(* Logix 5000 project; controller TFF vendor 1 type 14 code 107 rev 33.11; software revision 33.04; part 5 of 38 *)

        [0,11].PID.KP := 0.1, [0,11].PID.KI := 0.1, [0,11].PID.BIAS := 23.09767, [0,11].PID.DB := 0.001, [0,11].PID.MAXO := 100.0, [0,11].PID.UPD := 0.25, [0,11].PID.ERR := 0.20000005, [0,11].PID.MAXCV := 100.0, [0,11].PID.MAXTIE := 100.0, [0,11].PID.DATA[0] := -23.098158, [0,11].PID.DATA[3] := 0.20000005, [0,11].PID.DATA[4] := 0.20000005, [0,11].PID.DATA[5] := 0.024420025, [0,11].PID.DATA[6] := 1.0, [0,11].PID.DATA[7] := 4.0, [0,11].PID.DATA[8] := 0.1, [0,11].PID.DATA[9] := 0.1, [0,11].PID.DATA[11] := 0.1, [0,11].PID.DATA[12] := 0.1, [0,11].PID.DATA[15] := 1.0, [0,11].PID.DATA[16] := 1.0, [0,13].RampTimer.PRE := 3600000, [0,13].StableTimer.PRE := 2000, [0,13].PIDTimer.PRE := 10000, [0,13].PIDTimer.EN := 1, [0,13].PIDTimer.TT := 1, [0,13].PID.CTL := 305173120, [0,13].PID.PVT := 1, [0,13].PID.CA := 1, [0,13].PID.NOBC := 1, [0,13].PID.NOZC := 1, [0,13].PID.INI := 1, [0,13].PID.OLH := 1, [0,13].PID.DVPA := 1, [0,13].PID.PVHA := 1, [0,13].PID.KP := 0.2, [0,13].PID.KI := 0.08, [0,13].PID.MAXS := 100.0, [0,13].PID.DB := 1.0, [0,13].PID.SO := 100.0, [0,13].PID.MAXO := 100.0, [0,13].PID.UPD := 0.01, [0,13].PID.PV := 43.925232, [0,13].PID.ERR := 43.925232, [0,13].PID.OUT := 100.0, [0,13].PID.MAXI := 100.0, [0,13].PID.TIE := 2.4420025, [0,13].PID.MAXCV := 100.0, [0,13].PID.MAXTIE := 4095.0, [0,13].PID.DATA[0] := 100.0, [0,13].PID.DATA[1] := 702.8037, [0,13].PID.DATA[2] := 43.925232, [0,13].PID.DATA[3] := 43.925232, [0,13].PID.DATA[5] := 1.0, [0,13].PID.DATA[6] := 1.0, [0,13].PID.DATA[7] := 0.16, [0,13].PID.DATA[8] := 0.2, [0,13].PID.DATA[9] := 0.08, [0,13].PID.DATA[11] := 0.2, [0,13].PID.DATA[12] := 0.08,
        [0,13].PID.DATA[15] := 1.0, [0,13].PID.DATA[16] := 0.024420025, [1,0].RampTimer.PRE := 3600000, [1,0].StableTimer.PRE := 5000, [1,0].PIDTimer.PRE := 250, [1,0].PIDTimer.ACC := 100, [1,0].PIDTimer.EN := 1, [1,0].PIDTimer.TT := 1, [1,0].PID.CTL := 25199488, [1,0].PID.MO := 1, [1,0].PID.PE := 1, [1,0].PID.INI := 1, [1,0].PID.DVPA := 1, [1,0].PID.PVLA := 1, [1,0].PID.PVHA := 1, [1,0].PID.SP := 66.66666, [1,0].PID.KP := 0.5, [1,0].PID.KI := 0.1, [1,0].PID.MAXS := 200.0, [1,0].PID.SO := 10.0, [1,0].PID.MAXO := 100.0, [1,0].PID.MINO := 10.0, [1,0].PID.UPD := 0.25, [1,0].PID.ERR := 66.66666, [1,0].PID.OUT := 10.0, [1,0].PID.MAXI := 200.0, [1,0].PID.TIE := 10.0, [1,0].PID.MAXCV := 100.0, [1,0].PID.MAXTIE := 100.0, [1,0].PID.DATA[0] := -6.666666, [1,0].PID.DATA[3] := 66.66666, [1,0].PID.DATA[4] := 66.66666, [1,0].PID.DATA[5] := 0.5, [1,0].PID.DATA[6] := 1.0, [1,0].PID.DATA[7] := 4.0, [1,0].PID.DATA[8] := 0.5, [1,0].PID.DATA[9] := 0.1, [1,0].PID.DATA[11] := 0.5, [1,0].PID.DATA[12] := 0.08333334, [1,0].PID.DATA[15] := 1.0, [1,0].PID.DATA[16] := 1.0, [1,1].Tag := 'FIC01', [1,1].Desc := 'Prim. Feed Pump Control', [1,1].LoopCfg := 1, [1,1].ManualEGU := '%', [1,1].Auto1EGU := 'LPM', [1,1].Auto2EGU := 'cm/h', [1,1].Manual := 1, [1,1].DBOK := 1, [1,1].RampEnable := 1, [1,1].PIDEnable := 1, [1,1].ManualOSR := 1, [1,1].RangeMax := 100.0, [1,1].RampRate := 5.0, [1,1].RampRateSave := 5.0, [1,1].Deadband := 5.0, [1,1].RampTimer.PRE := 3600000, [1,1].StableTimer.PRE := 10000, [1,1].StableTime := 10, [1,1].PIDTimer.PRE := 250,
        [1,1].CycleTimer.PRE := 2000, [1,1].PID.CTL := -2080340096, [1,1].PID.EN := 1, [1,1].PID.SWM := 1, [1,1].PID.INI := 1, [1,1].PID.DVNA := 1, [1,1].PID.DVPA := 1, [1,1].PID.PVLA := 1, [1,1].PID.PVHA := 1, [1,1].PID.KP := 0.7, [1,1].PID.KI := 1.4, [1,1].PID.KD := 0.013, [1,1].PID.MAXS := 22.0, [1,1].PID.DB := 0.001, [1,1].PID.MAXO := 100.0, [1,1].PID.UPD := 0.25, [1,1].PID.MAXI := 22.0, [1,1].PID.MAXCV := 100.0, [1,1].PID.MAXTIE := 22.0, [1,1].PID.DATA[5] := 4.5454545, [1,1].PID.DATA[6] := 1.0, [1,1].PID.DATA[7] := 4.013, [1,1].PID.DATA[8] := 0.7, [1,1].PID.DATA[9] := 1.4, [1,1].PID.DATA[10] := 0.013, [1,1].PID.DATA[11] := 0.7, [1,1].PID.DATA[12] := 1.4, [1,1].PID.DATA[13] := 0.013, [1,1].PID.DATA[15] := 1.0, [1,1].PID.DATA[16] := 4.5454545, [1,1].KP[0] := 700.0, [1,1].KI[0] := 1400.0, [1,1].KD[0] := 13.0, [1,1].Auto1Cfg := 1, [1,1].Auto2Cfg := 1, [1,1].Auto1PVCfg := 10, [1,1].Auto2PVCfg := 42, [1,1].Auto1RangeMax := 22.0, [1,1].Auto2RangeMax := 9999.0, [1,2].Tag := 'FIC02', [1,2].Desc := 'Sec. Feed Pump Control', [1,2].LoopCfg := 1, [1,2].ManualEGU := '%', [1,2].Auto1EGU := 'LPM', [1,2].Auto2EGU := 'cm/h', [1,2].Interlock := 1, [1,2].Manual := 1, [1,2].DBOK := 1, [1,2].RampEnable := 1, [1,2].PIDEnable := 1, [1,2].ManualOSR := 1, [1,2].RangeMax := 100.0, [1,2].RampRate := 5.0, [1,2].RampRateSave := 5.0, [1,2].Deadband := 5.0, [1,2].RampTimer.PRE := 3600000, [1,2].StableTimer.PRE := 10000, [1,2].StableTime := 10, [1,2].PIDTimer.PRE := 250, [1,2].CycleTimer.PRE := 2000,
        [1,2].PID.CTL := -2080340096, [1,2].PID.EN := 1, [1,2].PID.SWM := 1, [1,2].PID.INI := 1, [1,2].PID.DVNA := 1, [1,2].PID.DVPA := 1, [1,2].PID.PVLA := 1, [1,2].PID.PVHA := 1, [1,2].PID.KP := 0.7, [1,2].PID.KI := 1.4, [1,2].PID.KD := 0.013, [1,2].PID.MAXS := 22.0, [1,2].PID.DB := 0.001, [1,2].PID.MAXO := 100.0, [1,2].PID.UPD := 0.25, [1,2].PID.MAXI := 22.0, [1,2].PID.MAXCV := 100.0, [1,2].PID.MAXTIE := 100.0, [1,2].PID.DATA[5] := 4.5454545, [1,2].PID.DATA[6] := 1.0, [1,2].PID.DATA[7] := 4.013, [1,2].PID.DATA[8] := 0.7, [1,2].PID.DATA[9] := 1.4, [1,2].PID.DATA[10] := 0.013, [1,2].PID.DATA[11] := 0.7, [1,2].PID.DATA[12] := 1.4, [1,2].PID.DATA[13] := 0.013, [1,2].PID.DATA[15] := 1.0, [1,2].PID.DATA[16] := 1.0, [1,2].KP[0] := 700.0, [1,2].KI[0] := 1400.0, [1,2].KD[0] := 13.0, [1,2].DisOSR := 1, [1,2].Auto1Cfg := 1, [1,2].Auto2Cfg := 1, [1,2].Auto1PVCfg := 12, [1,2].Auto2PVCfg := 43, [1,2].Auto1RangeMax := 22.0, [1,2].Auto2RangeMax := 9999.0, [1,2].OutputAddress := 1, [1,3].Tag := 'PCV12', [1,3].Desc := 'Post Column PCV012 Control', [1,3].LoopCfg := 1, [1,3].ManualEGU := '%', [1,3].Enable := 1, [1,3].Manual := 1, [1,3].Stable := 1, [1,3].DBOK := 1, [1,3].Status := 3, [1,3].RampEnable := 1, [1,3].PIDEnable := 1, [1,3].ManualOSR := 1, [1,3].RangeMax := 100.0, [1,3].RampRate := 5.0, [1,3].RampRateSave := 5.0, [1,3].RampStart := 20.0, [1,3].RampTimer.PRE := 3600000, [1,3].StableTimer.PRE := 2300, [1,3].StableTimer.ACC := 2354, [1,3].StableTimer.EN := 1,
        [1,3].StableTimer.DN := 1, [1,3].PIDTimer.PRE := 250, [1,3].CycleTimer.PRE := 2000, [1,3].PID.CTL := -1946122368, [1,3].PID.EN := 1, [1,3].PID.DOE := 1, [1,3].PID.SWM := 1, [1,3].PID.INI := 1, [1,3].PID.DVNA := 1, [1,3].PID.DVPA := 1, [1,3].PID.PVLA := 1, [1,3].PID.PVHA := 1, [1,3].PID.KP := 0.001, [1,3].PID.KI := 0.001, [1,3].PID.BIAS := 30.796, [1,3].PID.MAXS := 4095.0, [1,3].PID.MAXO := 100.0, [1,3].PID.UPD := 0.01, [1,3].PID.MAXI := 4095.0, [1,3].PID.MAXCV := 100.0, [1,3].PID.MAXTIE := 100.0, [1,3].PID.DATA[0] := -30.796, [1,3].PID.DATA[5] := 0.024420025, [1,3].PID.DATA[6] := 1.0, [1,3].PID.DATA[7] := 0.16, [1,3].PID.DATA[8] := 0.001, [1,3].PID.DATA[9] := 0.001, [1,3].PID.DATA[11] := 0.001, [1,3].PID.DATA[12] := 0.001, [1,3].PID.DATA[15] := 1.0, [1,3].PID.DATA[16] := 1.0, [1,3].OutputAddress := 2, [1,4].Tag := 'PCV10', [1,4].Desc := 'Line Pump1 PCV010 Control', [1,4].ManualEGU := '%', [1,4].Manual := 1, [1,4].Status := 3, [1,4].RampEnable := 1, [1,4].PIDEnable := 1, [1,4].RangeMax := 100.0, [1,4].RampRate := 0.5, [1,4].RampRateSave := 0.5, [1,4].RampStart := 3.443, [1,4].RampTimer.PRE := 3600000, [1,4].StableTimer.PRE := 5000, [1,4].PIDTimer.PRE := 250, [1,4].CycleTimer.PRE := 2000, [1,4].PID.CTL := 35652992, [1,4].PID.CA := 1, [1,4].PID.NOBC := 1, [1,4].PID.DVNA := 1, [1,4].PID.PVLA := 1, [1,4].PID.PVHA := 1, [1,4].PID.SP := 19.6, [1,4].PID.KP := 0.1, [1,4].PID.KI := 0.3, [1,4].PID.MAXS := 150.0, [1,4].PID.MAXO := 100.0, [1,4].PID.UPD := 0.25, [1,4].PID.ERR := -19.6,
        [1,4].PID.MAXI := 150.0, [1,4].PID.MAXCV := 100.0, [1,4].PID.MAXTIE := 100.0, [1,4].PID.DATA[0] := 1.3066667, [1,4].PID.DATA[3] := -19.6, [1,4].PID.DATA[4] := 19.6, [1,4].PID.DATA[5] := 0.6666667, [1,4].PID.DATA[6] := 1.0, [1,4].PID.DATA[7] := 4.0, [1,4].PID.DATA[8] := 0.1, [1,4].PID.DATA[9] := 0.3, [1,4].PID.DATA[11] := 0.1, [1,4].PID.DATA[12] := 0.3, [1,4].PID.DATA[15] := 1.0, [1,4].PID.DATA[16] := 1.0, [1,4].OutputAddress := 2, [1,5].Tag := 'PCV11', [1,5].Desc := 'Line Pump2 PCV011 Control', [1,5].ManualEGU := '%', [1,5].Manual := 1, [1,5].Status := 3, [1,5].RampEnable := 1, [1,5].PIDEnable := 1, [1,5].RangeMax := 100.0, [1,5].RampRate := 0.5, [1,5].RampRateSave := 0.5, [1,5].RampStart := 4.417, [1,5].RampTimer.PRE := 3600000, [1,5].StableTimer.PRE := 1500, [1,5].PIDTimer.PRE := 250, [1,5].CycleTimer.PRE := 2000, [1,5].PID.CTL := 134218624, [1,5].PID.DOE := 1, [1,5].PID.DVPA := 1, [1,5].PID.PVLA := 1, [1,5].PID.PVHA := 1, [1,5].PID.SP := 350.0, [1,5].PID.KP := 40.0, [1,5].PID.KI := 0.5, [1,5].PID.BIAS := -847.4798, [1,5].PID.MAXS := 550.0, [1,5].PID.MAXO := 100.0, [1,5].PID.UPD := 0.25, [1,5].PID.ERR := 350.0, [1,5].PID.MAXI := 550.0, [1,5].PID.MAXCV := 100.0, [1,5].PID.MAXTIE := 100.0, [1,5].PID.DATA[0] := -1697.9749, [1,5].PID.DATA[1] := 1018.1818, [1,5].PID.DATA[3] := 350.0, [1,5].PID.DATA[4] := 350.0, [1,5].PID.DATA[5] := 0.18181819, [1,5].PID.DATA[6] := 1.0, [1,5].PID.DATA[7] := 4.0, [1,5].PID.DATA[8] := 40.0, [1,5].PID.DATA[9] := 0.5, [1,5].PID.DATA[11] := 40.0, [1,5].PID.DATA[12] := 0.5, [1,5].PID.DATA[15] := 1.0, [1,5].PID.DATA[16] := 1.0,
        [1,5].OutputAddress := 3, [1,6].StableTimer.PRE := 15000, [1,6].PIDTimer.EN := 1, [1,6].PIDTimer.TT := 1, [1,6].CycleTimer.PRE := 5000, [1,6].PID.CTL := 16810624, [1,6].PID.MO := 1, [1,6].PID.INI := 1, [1,6].PID.DVPA := 1, [1,6].PID.PVHA := 1, [1,6].PID.SP := 10.0, [1,6].PID.KP := 0.3, [1,6].PID.KI := 0.3, [1,6].PID.MAXS := 200.0, [1,6].PID.SO := 3.074094, [1,6].PID.MAXO := 100.0, [1,6].PID.UPD := 0.25, [1,6].PID.PV := 1.488363, [1,6].PID.ERR := 8.511638, [1,6].PID.OUT := 3.074094, [1,6].PID.MAXI := 200.0, [1,6].PID.TIE := 3.074094, [1,6].PID.MAXCV := 200.0, [1,6].PID.MAXTIE := 200.0, [1,6].PID.DATA[0] := 1.797348, [1,6].PID.DATA[1] := -11.9069, [1,6].PID.DATA[2] := 1.488363, [1,6].PID.DATA[3] := 8.511638, [1,6].PID.DATA[4] := 10.0, [1,6].PID.DATA[5] := 0.5, [1,6].PID.DATA[6] := 1.0, [1,6].PID.DATA[7] := 4.0, [1,6].PID.DATA[8] := 0.3, [1,6].PID.DATA[9] := 0.3, [1,6].PID.DATA[11] := 0.3, [1,6].PID.DATA[12] := 0.3, [1,6].PID.DATA[15] := 2.0, [1,6].PID.DATA[16] := 0.5, [1,7].StableTimer.PRE := 200, [1,7].PIDTimer.PRE := 250, [1,7].PIDTimer.EN := 1, [1,7].PIDTimer.TT := 1, [1,7].CycleTimer.PRE := 10000, [1,7].PID.CTL := 16810880, [1,7].PID.MO := 1, [1,7].PID.INI := 1, [1,7].PID.DVPA := 1, [1,7].PID.PVLA := 1, [1,7].PID.PVHA := 1, [1,7].PID.SP := 10.0, [1,7].PID.KP := 2.0, [1,7].PID.KI := 0.2, [1,7].PID.KD := 0.3, [1,7].PID.BIAS := 50.0, [1,7].PID.DB := 0.01, [1,7].PID.SO := 80.0, [1,7].PID.MAXO := 100.0, [1,7].PID.UPD := 0.25, [1,7].PID.ERR := 10.0, [1,7].PID.OUT := 80.0,
        [1,7].PID.TIE := 80.0, [1,7].PID.MAXCV := 100.0, [1,7].PID.MAXTIE := 100.0, [1,7].PID.DATA[0] := 29.511597, [1,7].PID.DATA[3] := 10.0, [1,7].PID.DATA[4] := 10.0, [1,7].PID.DATA[5] := 0.024420025, [1,7].PID.DATA[6] := 1.0, [1,7].PID.DATA[7] := 4.3, [1,7].PID.DATA[8] := 2.0, [1,7].PID.DATA[9] := 0.2, [1,7].PID.DATA[10] := 0.3, [1,7].PID.DATA[11] := 2.0, [1,7].PID.DATA[12] := 0.2, [1,7].PID.DATA[13] := 0.3, [1,7].PID.DATA[15] := 1.0, [1,7].PID.DATA[16] := 1.0, [1,8].StableTimer.PRE := 15000, [1,8].PIDTimer.PRE := 250, [1,8].CycleTimer.PRE := 20000, [1,8].PID.CTL := 33555584, [1,8].PID.CA := 1, [1,8].PID.DVNA := 1, [1,8].PID.PVHA := 1, [1,8].PID.SP := 27.0, [1,8].PID.KP := 1.0, [1,8].PID.KI := 0.1, [1,8].PID.MAXS := 100.0, [1,8].PID.MAXO := 100.0, [1,8].PID.UPD := 0.25, [1,8].PID.PV := 18.2328, [1,8].PID.ERR := -8.767202, [1,8].PID.MAXI := 100.0, [1,8].PID.MAXCV := 100.0, [1,8].PID.MAXTIE := 100.0, [1,8].PID.DATA[0] := 8.767202, [1,8].PID.DATA[1] := 291.7248, [1,8].PID.DATA[2] := 18.2328, [1,8].PID.DATA[3] := -8.767202, [1,8].PID.DATA[4] := 27.0, [1,8].PID.DATA[5] := 1.0, [1,8].PID.DATA[6] := 1.0, [1,8].PID.DATA[7] := 4.0, [1,8].PID.DATA[8] := 1.0, [1,8].PID.DATA[9] := 0.1, [1,8].PID.DATA[11] := 1.0, [1,8].PID.DATA[12] := 0.1, [1,8].PID.DATA[15] := 1.0, [1,8].PID.DATA[16] := 1.0, [1,11].RampTimer.PRE := 100000, [1,11].StableTimer.PRE := 200, [1,11].PIDTimer.PRE := 250, [1,11].PIDTimer.ACC := 230, [1,11].PIDTimer.EN := 1, [1,11].PIDTimer.TT := 1, [1,11].PID.CTL := 67142528, [1,11].PID.SWM := 1, [1,11].PID.INI := 1, [1,11].PID.DVPA := 1, [1,11].PID.PVLA := 1,
        [1,11].PID.PVHA := 1, [1,11].PID.SP := 0.20000005, [1,11].PID.KP := 0.1, [1,11].PID.KI := 0.1, [1,11].PID.BIAS := 23.09767, [1,11].PID.DB := 0.001, [1,11].PID.MAXO := 100.0, [1,11].PID.UPD := 0.25, [1,11].PID.ERR := 0.20000005, [1,11].PID.MAXCV := 100.0, [1,11].PID.MAXTIE := 100.0, [1,11].PID.DATA[0] := -23.098158, [1,11].PID.DATA[3] := 0.20000005, [1,11].PID.DATA[4] := 0.20000005, [1,11].PID.DATA[5] := 0.024420025, [1,11].PID.DATA[6] := 1.0, [1,11].PID.DATA[7] := 4.0, [1,11].PID.DATA[8] := 0.1, [1,11].PID.DATA[9] := 0.1, [1,11].PID.DATA[11] := 0.1, [1,11].PID.DATA[12] := 0.1, [1,11].PID.DATA[15] := 1.0, [1,11].PID.DATA[16] := 1.0, [1,13].RampTimer.PRE := 3600000, [1,13].StableTimer.PRE := 2000, [1,13].PIDTimer.PRE := 10000, [1,13].PIDTimer.EN := 1, [1,13].PIDTimer.TT := 1, [1,13].PID.CTL := 305173120, [1,13].PID.PVT := 1, [1,13].PID.CA := 1, [1,13].PID.NOBC := 1, [1,13].PID.NOZC := 1, [1,13].PID.INI := 1, [1,13].PID.OLH := 1, [1,13].PID.DVPA := 1, [1,13].PID.PVHA := 1, [1,13].PID.KP := 0.2, [1,13].PID.KI := 0.08, [1,13].PID.MAXS := 100.0, [1,13].PID.DB := 1.0, [1,13].PID.SO := 100.0, [1,13].PID.MAXO := 100.0, [1,13].PID.UPD := 0.01, [1,13].PID.PV := 43.925232, [1,13].PID.ERR := 43.925232, [1,13].PID.OUT := 100.0, [1,13].PID.MAXI := 100.0, [1,13].PID.TIE := 2.4420025, [1,13].PID.MAXCV := 100.0, [1,13].PID.MAXTIE := 4095.0, [1,13].PID.DATA[0] := 100.0, [1,13].PID.DATA[1] := 702.8037, [1,13].PID.DATA[2] := 43.925232, [1,13].PID.DATA[3] := 43.925232, [1,13].PID.DATA[5] := 1.0, [1,13].PID.DATA[6] := 1.0, [1,13].PID.DATA[7] := 0.16, [1,13].PID.DATA[8] := 0.2, [1,13].PID.DATA[9] := 0.08,
        [1,13].PID.DATA[11] := 0.2, [1,13].PID.DATA[12] := 0.08, [1,13].PID.DATA[15] := 1.0, [1,13].PID.DATA[16] := 0.024420025, [2,0].RampTimer.PRE := 3600000, [2,0].StableTimer.PRE := 5000, [2,0].PIDTimer.PRE := 250, [2,0].PIDTimer.ACC := 100, [2,0].PIDTimer.EN := 1, [2,0].PIDTimer.TT := 1, [2,0].PID.CTL := 25199488, [2,0].PID.MO := 1, [2,0].PID.PE := 1, [2,0].PID.INI := 1, [2,0].PID.DVPA := 1, [2,0].PID.PVLA := 1, [2,0].PID.PVHA := 1, [2,0].PID.SP := 66.66666, [2,0].PID.KP := 0.5, [2,0].PID.KI := 0.1, [2,0].PID.MAXS := 200.0, [2,0].PID.SO := 10.0, [2,0].PID.MAXO := 100.0, [2,0].PID.MINO := 10.0, [2,0].PID.UPD := 0.25, [2,0].PID.ERR := 66.66666, [2,0].PID.OUT := 10.0, [2,0].PID.MAXI := 200.0, [2,0].PID.TIE := 10.0, [2,0].PID.MAXCV := 100.0, [2,0].PID.MAXTIE := 100.0, [2,0].PID.DATA[0] := -6.666666, [2,0].PID.DATA[3] := 66.66666, [2,0].PID.DATA[4] := 66.66666, [2,0].PID.DATA[5] := 0.5, [2,0].PID.DATA[6] := 1.0, [2,0].PID.DATA[7] := 4.0, [2,0].PID.DATA[8] := 0.5, [2,0].PID.DATA[9] := 0.1, [2,0].PID.DATA[11] := 0.5, [2,0].PID.DATA[12] := 0.08333334, [2,0].PID.DATA[15] := 1.0, [2,0].PID.DATA[16] := 1.0, [2,1].Tag := 'FIC01', [2,1].Desc := 'Prim. Feed Pump Control', [2,1].LoopCfg := 1, [2,1].ManualEGU := '%', [2,1].Auto1EGU := 'LPM', [2,1].Auto2EGU := 'cm/h', [2,1].Manual := 1, [2,1].DBOK := 1, [2,1].RampEnable := 1, [2,1].PIDEnable := 1, [2,1].ManualOSR := 1, [2,1].RangeMax := 100.0, [2,1].RampRate := 5.0, [2,1].RampRateSave := 5.0, [2,1].Deadband := 5.0, [2,1].RampTimer.PRE := 3600000, [2,1].StableTimer.PRE := 10000,
        [2,1].StableTime := 10, [2,1].PIDTimer.PRE := 250, [2,1].CycleTimer.PRE := 2000, [2,1].PID.CTL := -2080340096, [2,1].PID.EN := 1, [2,1].PID.SWM := 1, [2,1].PID.INI := 1, [2,1].PID.DVNA := 1, [2,1].PID.DVPA := 1, [2,1].PID.PVLA := 1, [2,1].PID.PVHA := 1, [2,1].PID.KP := 0.7, [2,1].PID.KI := 1.4, [2,1].PID.KD := 0.013, [2,1].PID.MAXS := 22.0, [2,1].PID.DB := 0.001, [2,1].PID.MAXO := 100.0, [2,1].PID.UPD := 0.25, [2,1].PID.MAXI := 22.0, [2,1].PID.MAXCV := 100.0, [2,1].PID.MAXTIE := 22.0, [2,1].PID.DATA[5] := 4.5454545, [2,1].PID.DATA[6] := 1.0, [2,1].PID.DATA[7] := 4.013, [2,1].PID.DATA[8] := 0.7, [2,1].PID.DATA[9] := 1.4, [2,1].PID.DATA[10] := 0.013, [2,1].PID.DATA[11] := 0.7, [2,1].PID.DATA[12] := 1.4, [2,1].PID.DATA[13] := 0.013, [2,1].PID.DATA[15] := 1.0, [2,1].PID.DATA[16] := 4.5454545, [2,1].KP[0] := 700.0, [2,1].KI[0] := 1400.0, [2,1].KD[0] := 13.0, [2,1].Auto1Cfg := 1, [2,1].Auto2Cfg := 1, [2,1].Auto1PVCfg := 10, [2,1].Auto2PVCfg := 42, [2,1].Auto1RangeMax := 22.0, [2,1].Auto2RangeMax := 9999.0, [2,2].Tag := 'FIC02', [2,2].Desc := 'Sec. Feed Pump Control', [2,2].LoopCfg := 1, [2,2].ManualEGU := '%', [2,2].Auto1EGU := 'LPM', [2,2].Auto2EGU := 'cm/h', [2,2].Interlock := 1, [2,2].Manual := 1, [2,2].DBOK := 1, [2,2].RampEnable := 1, [2,2].PIDEnable := 1, [2,2].ManualOSR := 1, [2,2].RangeMax := 100.0, [2,2].RampRate := 5.0, [2,2].RampRateSave := 5.0, [2,2].Deadband := 5.0, [2,2].RampTimer.PRE := 3600000, [2,2].StableTimer.PRE := 10000, [2,2].StableTime := 10,
        [2,2].PIDTimer.PRE := 250, [2,2].CycleTimer.PRE := 2000, [2,2].PID.CTL := -2080340096, [2,2].PID.EN := 1, [2,2].PID.SWM := 1, [2,2].PID.INI := 1, [2,2].PID.DVNA := 1, [2,2].PID.DVPA := 1, [2,2].PID.PVLA := 1, [2,2].PID.PVHA := 1, [2,2].PID.KP := 0.7, [2,2].PID.KI := 1.4, [2,2].PID.KD := 0.013, [2,2].PID.MAXS := 22.0, [2,2].PID.DB := 0.001, [2,2].PID.MAXO := 100.0, [2,2].PID.UPD := 0.25, [2,2].PID.MAXI := 22.0, [2,2].PID.MAXCV := 100.0, [2,2].PID.MAXTIE := 100.0, [2,2].PID.DATA[5] := 4.5454545, [2,2].PID.DATA[6] := 1.0, [2,2].PID.DATA[7] := 4.013, [2,2].PID.DATA[8] := 0.7, [2,2].PID.DATA[9] := 1.4, [2,2].PID.DATA[10] := 0.013, [2,2].PID.DATA[11] := 0.7, [2,2].PID.DATA[12] := 1.4, [2,2].PID.DATA[13] := 0.013, [2,2].PID.DATA[15] := 1.0, [2,2].PID.DATA[16] := 1.0, [2,2].KP[0] := 700.0, [2,2].KI[0] := 1400.0, [2,2].KD[0] := 13.0, [2,2].DisOSR := 1, [2,2].Auto1Cfg := 1, [2,2].Auto2Cfg := 1, [2,2].Auto1PVCfg := 12, [2,2].Auto2PVCfg := 43, [2,2].Auto1RangeMax := 22.0, [2,2].Auto2RangeMax := 9999.0, [2,2].OutputAddress := 1, [2,3].Tag := 'PCV12', [2,3].Desc := 'Post Column PCV012 Control', [2,3].LoopCfg := 1, [2,3].ManualEGU := '%', [2,3].Enable := 1, [2,3].Manual := 1, [2,3].Stable := 1, [2,3].DBOK := 1, [2,3].Status := 3, [2,3].RampEnable := 1, [2,3].PIDEnable := 1, [2,3].ManualOSR := 1, [2,3].RangeMax := 100.0, [2,3].RampRate := 5.0, [2,3].RampRateSave := 5.0, [2,3].RampStart := 20.0, [2,3].RampTimer.PRE := 3600000, [2,3].StableTimer.PRE := 2300,
        [2,3].StableTimer.ACC := 2354, [2,3].StableTimer.EN := 1, [2,3].StableTimer.DN := 1, [2,3].PIDTimer.PRE := 250, [2,3].CycleTimer.PRE := 2000, [2,3].PID.CTL := -1946122368, [2,3].PID.EN := 1, [2,3].PID.DOE := 1, [2,3].PID.SWM := 1, [2,3].PID.INI := 1, [2,3].PID.DVNA := 1, [2,3].PID.DVPA := 1, [2,3].PID.PVLA := 1, [2,3].PID.PVHA := 1, [2,3].PID.KP := 0.001, [2,3].PID.KI := 0.001, [2,3].PID.BIAS := 30.796, [2,3].PID.MAXS := 4095.0, [2,3].PID.MAXO := 100.0, [2,3].PID.UPD := 0.01, [2,3].PID.MAXI := 4095.0, [2,3].PID.MAXCV := 100.0, [2,3].PID.MAXTIE := 100.0, [2,3].PID.DATA[0] := -30.796, [2,3].PID.DATA[5] := 0.024420025, [2,3].PID.DATA[6] := 1.0, [2,3].PID.DATA[7] := 0.16, [2,3].PID.DATA[8] := 0.001, [2,3].PID.DATA[9] := 0.001, [2,3].PID.DATA[11] := 0.001, [2,3].PID.DATA[12] := 0.001, [2,3].PID.DATA[15] := 1.0, [2,3].PID.DATA[16] := 1.0, [2,3].OutputAddress := 2, [2,4].Tag := 'PCV10', [2,4].Desc := 'Line Pump1 PCV010 Control', [2,4].ManualEGU := '%', [2,4].Manual := 1, [2,4].Status := 3, [2,4].RampEnable := 1, [2,4].PIDEnable := 1, [2,4].RangeMax := 100.0, [2,4].RampRate := 0.5, [2,4].RampRateSave := 0.5, [2,4].RampStart := 3.443, [2,4].RampTimer.PRE := 3600000, [2,4].StableTimer.PRE := 5000, [2,4].PIDTimer.PRE := 250, [2,4].CycleTimer.PRE := 2000, [2,4].PID.CTL := 35652992, [2,4].PID.CA := 1, [2,4].PID.NOBC := 1, [2,4].PID.DVNA := 1, [2,4].PID.PVLA := 1, [2,4].PID.PVHA := 1, [2,4].PID.SP := 19.6, [2,4].PID.KP := 0.1, [2,4].PID.KI := 0.3, [2,4].PID.MAXS := 150.0, [2,4].PID.MAXO := 100.0,
        [2,4].PID.UPD := 0.25, [2,4].PID.ERR := -19.6, [2,4].PID.MAXI := 150.0, [2,4].PID.MAXCV := 100.0, [2,4].PID.MAXTIE := 100.0, [2,4].PID.DATA[0] := 1.3066667, [2,4].PID.DATA[3] := -19.6, [2,4].PID.DATA[4] := 19.6, [2,4].PID.DATA[5] := 0.6666667, [2,4].PID.DATA[6] := 1.0, [2,4].PID.DATA[7] := 4.0, [2,4].PID.DATA[8] := 0.1, [2,4].PID.DATA[9] := 0.3, [2,4].PID.DATA[11] := 0.1, [2,4].PID.DATA[12] := 0.3, [2,4].PID.DATA[15] := 1.0, [2,4].PID.DATA[16] := 1.0, [2,4].OutputAddress := 2, [2,5].Tag := 'PCV11', [2,5].Desc := 'Line Pump2 PCV011 Control', [2,5].ManualEGU := '%', [2,5].Manual := 1, [2,5].Status := 3, [2,5].RampEnable := 1, [2,5].PIDEnable := 1, [2,5].RangeMax := 100.0, [2,5].RampRate := 0.5, [2,5].RampRateSave := 0.5, [2,5].RampStart := 4.417, [2,5].RampTimer.PRE := 3600000, [2,5].StableTimer.PRE := 1500, [2,5].PIDTimer.PRE := 250, [2,5].CycleTimer.PRE := 2000, [2,5].PID.CTL := 134218624, [2,5].PID.DOE := 1, [2,5].PID.DVPA := 1, [2,5].PID.PVLA := 1, [2,5].PID.PVHA := 1, [2,5].PID.SP := 350.0, [2,5].PID.KP := 40.0, [2,5].PID.KI := 0.5, [2,5].PID.BIAS := -847.4798, [2,5].PID.MAXS := 550.0, [2,5].PID.MAXO := 100.0, [2,5].PID.UPD := 0.25, [2,5].PID.ERR := 350.0, [2,5].PID.MAXI := 550.0, [2,5].PID.MAXCV := 100.0, [2,5].PID.MAXTIE := 100.0, [2,5].PID.DATA[0] := -1697.9749, [2,5].PID.DATA[1] := 1018.1818, [2,5].PID.DATA[3] := 350.0, [2,5].PID.DATA[4] := 350.0, [2,5].PID.DATA[5] := 0.18181819, [2,5].PID.DATA[6] := 1.0, [2,5].PID.DATA[7] := 4.0, [2,5].PID.DATA[8] := 40.0, [2,5].PID.DATA[9] := 0.5, [2,5].PID.DATA[11] := 40.0, [2,5].PID.DATA[12] := 0.5,
        [2,5].PID.DATA[15] := 1.0, [2,5].PID.DATA[16] := 1.0, [2,5].OutputAddress := 3, [2,6].StableTimer.PRE := 15000, [2,6].PIDTimer.EN := 1, [2,6].PIDTimer.TT := 1, [2,6].CycleTimer.PRE := 5000, [2,6].PID.CTL := 16810624, [2,6].PID.MO := 1, [2,6].PID.INI := 1, [2,6].PID.DVPA := 1, [2,6].PID.PVHA := 1, [2,6].PID.SP := 10.0, [2,6].PID.KP := 0.3, [2,6].PID.KI := 0.3, [2,6].PID.MAXS := 200.0, [2,6].PID.SO := 3.074094, [2,6].PID.MAXO := 100.0, [2,6].PID.UPD := 0.25, [2,6].PID.PV := 1.488363, [2,6].PID.ERR := 8.511638, [2,6].PID.OUT := 3.074094, [2,6].PID.MAXI := 200.0, [2,6].PID.TIE := 3.074094, [2,6].PID.MAXCV := 200.0, [2,6].PID.MAXTIE := 200.0, [2,6].PID.DATA[0] := 1.797348, [2,6].PID.DATA[1] := -11.9069, [2,6].PID.DATA[2] := 1.488363, [2,6].PID.DATA[3] := 8.511638, [2,6].PID.DATA[4] := 10.0, [2,6].PID.DATA[5] := 0.5, [2,6].PID.DATA[6] := 1.0, [2,6].PID.DATA[7] := 4.0, [2,6].PID.DATA[8] := 0.3, [2,6].PID.DATA[9] := 0.3, [2,6].PID.DATA[11] := 0.3, [2,6].PID.DATA[12] := 0.3, [2,6].PID.DATA[15] := 2.0, [2,6].PID.DATA[16] := 0.5, [2,7].StableTimer.PRE := 200, [2,7].PIDTimer.PRE := 250, [2,7].PIDTimer.EN := 1, [2,7].PIDTimer.TT := 1, [2,7].CycleTimer.PRE := 10000, [2,7].PID.CTL := 16810880, [2,7].PID.MO := 1, [2,7].PID.INI := 1, [2,7].PID.DVPA := 1, [2,7].PID.PVLA := 1, [2,7].PID.PVHA := 1, [2,7].PID.SP := 10.0, [2,7].PID.KP := 2.0, [2,7].PID.KI := 0.2, [2,7].PID.KD := 0.3, [2,7].PID.BIAS := 50.0, [2,7].PID.DB := 0.01, [2,7].PID.SO := 80.0, [2,7].PID.MAXO := 100.0, [2,7].PID.UPD := 0.25,
        [2,7].PID.ERR := 10.0, [2,7].PID.OUT := 80.0, [2,7].PID.TIE := 80.0, [2,7].PID.MAXCV := 100.0, [2,7].PID.MAXTIE := 100.0, [2,7].PID.DATA[0] := 29.511597, [2,7].PID.DATA[3] := 10.0, [2,7].PID.DATA[4] := 10.0, [2,7].PID.DATA[5] := 0.024420025, [2,7].PID.DATA[6] := 1.0, [2,7].PID.DATA[7] := 4.3, [2,7].PID.DATA[8] := 2.0, [2,7].PID.DATA[9] := 0.2, [2,7].PID.DATA[10] := 0.3, [2,7].PID.DATA[11] := 2.0, [2,7].PID.DATA[12] := 0.2, [2,7].PID.DATA[13] := 0.3, [2,7].PID.DATA[15] := 1.0, [2,7].PID.DATA[16] := 1.0, [2,8].StableTimer.PRE := 15000, [2,8].PIDTimer.PRE := 250, [2,8].CycleTimer.PRE := 20000, [2,8].PID.CTL := 33555584, [2,8].PID.CA := 1, [2,8].PID.DVNA := 1, [2,8].PID.PVHA := 1, [2,8].PID.SP := 27.0, [2,8].PID.KP := 1.0, [2,8].PID.KI := 0.1, [2,8].PID.MAXS := 100.0, [2,8].PID.MAXO := 100.0, [2,8].PID.UPD := 0.25, [2,8].PID.PV := 18.2328, [2,8].PID.ERR := -8.767202, [2,8].PID.MAXI := 100.0, [2,8].PID.MAXCV := 100.0, [2,8].PID.MAXTIE := 100.0, [2,8].PID.DATA[0] := 8.767202, [2,8].PID.DATA[1] := 291.7248, [2,8].PID.DATA[2] := 18.2328, [2,8].PID.DATA[3] := -8.767202, [2,8].PID.DATA[4] := 27.0, [2,8].PID.DATA[5] := 1.0, [2,8].PID.DATA[6] := 1.0, [2,8].PID.DATA[7] := 4.0, [2,8].PID.DATA[8] := 1.0, [2,8].PID.DATA[9] := 0.1, [2,8].PID.DATA[11] := 1.0, [2,8].PID.DATA[12] := 0.1, [2,8].PID.DATA[15] := 1.0, [2,8].PID.DATA[16] := 1.0, [2,11].RampTimer.PRE := 100000, [2,11].StableTimer.PRE := 200, [2,11].PIDTimer.PRE := 250, [2,11].PIDTimer.ACC := 230, [2,11].PIDTimer.EN := 1, [2,11].PIDTimer.TT := 1, [2,11].PID.CTL := 67142528, [2,11].PID.SWM := 1, [2,11].PID.INI := 1,
        [2,11].PID.DVPA := 1, [2,11].PID.PVLA := 1, [2,11].PID.PVHA := 1, [2,11].PID.SP := 0.20000005, [2,11].PID.KP := 0.1, [2,11].PID.KI := 0.1, [2,11].PID.BIAS := 23.09767, [2,11].PID.DB := 0.001, [2,11].PID.MAXO := 100.0, [2,11].PID.UPD := 0.25, [2,11].PID.ERR := 0.20000005, [2,11].PID.MAXCV := 100.0, [2,11].PID.MAXTIE := 100.0, [2,11].PID.DATA[0] := -23.098158, [2,11].PID.DATA[3] := 0.20000005, [2,11].PID.DATA[4] := 0.20000005, [2,11].PID.DATA[5] := 0.024420025, [2,11].PID.DATA[6] := 1.0, [2,11].PID.DATA[7] := 4.0, [2,11].PID.DATA[8] := 0.1, [2,11].PID.DATA[9] := 0.1, [2,11].PID.DATA[11] := 0.1, [2,11].PID.DATA[12] := 0.1, [2,11].PID.DATA[15] := 1.0, [2,11].PID.DATA[16] := 1.0, [2,13].RampTimer.PRE := 3600000, [2,13].StableTimer.PRE := 2000, [2,13].PIDTimer.PRE := 10000, [2,13].PIDTimer.EN := 1, [2,13].PIDTimer.TT := 1, [2,13].PID.CTL := 305173120, [2,13].PID.PVT := 1, [2,13].PID.CA := 1, [2,13].PID.NOBC := 1, [2,13].PID.NOZC := 1, [2,13].PID.INI := 1, [2,13].PID.OLH := 1, [2,13].PID.DVPA := 1, [2,13].PID.PVHA := 1, [2,13].PID.KP := 0.2, [2,13].PID.KI := 0.08, [2,13].PID.MAXS := 100.0, [2,13].PID.DB := 1.0, [2,13].PID.SO := 100.0, [2,13].PID.MAXO := 100.0, [2,13].PID.UPD := 0.01, [2,13].PID.PV := 43.925232, [2,13].PID.ERR := 43.925232, [2,13].PID.OUT := 100.0, [2,13].PID.MAXI := 100.0, [2,13].PID.TIE := 2.4420025, [2,13].PID.MAXCV := 100.0, [2,13].PID.MAXTIE := 4095.0, [2,13].PID.DATA[0] := 100.0, [2,13].PID.DATA[1] := 702.8037, [2,13].PID.DATA[2] := 43.925232, [2,13].PID.DATA[3] := 43.925232, [2,13].PID.DATA[5] := 1.0, [2,13].PID.DATA[6] := 1.0, [2,13].PID.DATA[7] := 0.16,
        [2,13].PID.DATA[8] := 0.2, [2,13].PID.DATA[9] := 0.08, [2,13].PID.DATA[11] := 0.2, [2,13].PID.DATA[12] := 0.08, [2,13].PID.DATA[15] := 1.0, [2,13].PID.DATA[16] := 0.024420025, [3,1].LoopCfg := 1, [3,1].DBOK := 1, [3,1].RampEnable := 1, [3,1].PIDEnable := 1, [3,1].RangeMax := 100.0, [3,1].RampRate := 0.5, [3,1].RampRateSave := 0.5, [3,1].RampTimer.PRE := 3600000, [3,1].PIDTimer.PRE := 250, [3,1].PIDTimer.EN := 1, [3,1].PIDTimer.TT := 1, [3,1].CycleTimer.PRE := 2000, [3,1].PID.CTL := 67108864, [3,1].PID.SWM := 1, [3,1].PID.MAXS := 25.0, [3,1].PID.MAXO := 100.0, [3,1].PID.MAXI := 25.0, [3,1].PID.MAXCV := 100.0, [3,1].PID.MAXTIE := 25.0, [3,1].PID.DATA[5] := 4.0, [3,1].PID.DATA[6] := 1.0, [3,1].PID.DATA[15] := 1.0, [3,1].PID.DATA[16] := 4.0, [3,1].Auto1Cfg := 1, [3,1].Auto2Cfg := 1, [3,1].Auto1PVCfg := 10, [3,1].Auto2PVCfg := 42, [3,1].Auto1RangeMax := 55.0, [3,2].LoopCfg := 1, [3,2].DBOK := 1, [3,2].RampEnable := 1, [3,2].PIDEnable := 1, [3,2].RangeMax := 100.0, [3,2].RampRate := 0.5, [3,2].RampRateSave := 0.5, [3,2].RampTimer.PRE := 3600000, [3,2].PIDTimer.PRE := 250, [3,2].PIDTimer.EN := 1, [3,2].PIDTimer.TT := 1, [3,2].CycleTimer.PRE := 2000, [3,2].PID.CTL := 67108864, [3,2].PID.SWM := 1, [3,2].PID.MAXO := 100.0, [3,2].PID.MAXCV := 100.0, [3,2].PID.MAXTIE := 100.0, [3,2].PID.DATA[5] := 0.024420025, [3,2].PID.DATA[6] := 1.0, [3,2].PID.DATA[15] := 1.0, [3,2].PID.DATA[16] := 1.0, [3,2].Auto1Cfg := 1, [3,2].Auto2Cfg := 1, [3,2].Auto1PVCfg := 12, [3,2].Auto2PVCfg := 43, [3,2].Auto1RangeMax := 30.0,
        [3,2].OutputAddress := 1, [3,3].LoopCfg := 1, [3,3].Enable := 1, [3,3].Manual := 1, [3,3].Status := 9, [3,3].RampEnable := 1, [3,3].PIDEnable := 1, [3,3].RangeMax := 100.0, [3,3].RampRate := 0.5, [3,3].RampRateSave := 0.5, [3,3].RampTimer.PRE := 3600000, [3,3].PIDTimer.PRE := 250, [3,3].PIDTimer.EN := 1, [3,3].PIDTimer.TT := 1, [3,3].CycleTimer.PRE := 2000, [3,3].PID.CTL := 67108864, [3,3].PID.SWM := 1, [3,3].PID.MAXS := 4095.0, [3,3].PID.MAXO := 100.0, [3,3].PID.MAXI := 4095.0, [3,3].PID.MAXCV := 100.0, [3,3].PID.MAXTIE := 100.0, [3,3].PID.DATA[5] := 0.024420025, [3,3].PID.DATA[6] := 1.0, [3,3].PID.DATA[15] := 1.0, [3,3].PID.DATA[16] := 1.0, [3,3].OutputAddress := 2, [4,0].RampTimer.PRE := 3600000, [4,0].StableTimer.PRE := 5000, [4,0].PIDTimer.PRE := 250, [4,0].PIDTimer.ACC := 100, [4,0].PIDTimer.EN := 1, [4,0].PIDTimer.TT := 1, [4,0].PID.CTL := 25199488, [4,0].PID.MO := 1, [4,0].PID.PE := 1, [4,0].PID.INI := 1, [4,0].PID.DVPA := 1, [4,0].PID.PVLA := 1, [4,0].PID.PVHA := 1, [4,0].PID.SP := 66.66666, [4,0].PID.KP := 0.5, [4,0].PID.KI := 0.1, [4,0].PID.MAXS := 200.0, [4,0].PID.SO := 10.0, [4,0].PID.MAXO := 100.0, [4,0].PID.MINO := 10.0, [4,0].PID.UPD := 0.25, [4,0].PID.ERR := 66.66666, [4,0].PID.OUT := 10.0, [4,0].PID.MAXI := 200.0, [4,0].PID.TIE := 10.0, [4,0].PID.MAXCV := 100.0, [4,0].PID.MAXTIE := 100.0, [4,0].PID.DATA[0] := -6.666666, [4,0].PID.DATA[3] := 66.66666, [4,0].PID.DATA[4] := 66.66666, [4,0].PID.DATA[5] := 0.5, [4,0].PID.DATA[6] := 1.0, [4,0].PID.DATA[7] := 4.0,
        [4,0].PID.DATA[8] := 0.5, [4,0].PID.DATA[9] := 0.1, [4,0].PID.DATA[11] := 0.5, [4,0].PID.DATA[12] := 0.08333334, [4,0].PID.DATA[15] := 1.0, [4,0].PID.DATA[16] := 1.0, [4,1].Tag := 'FIC01', [4,1].Desc := 'Prim. Feed Pump Control', [4,1].LoopCfg := 1, [4,1].ManualEGU := '%', [4,1].Auto1EGU := 'LPM', [4,1].Auto2EGU := 'cm/h', [4,1].Manual := 1, [4,1].DBOK := 1, [4,1].RampEnable := 1, [4,1].PIDEnable := 1, [4,1].ManualOSR := 1, [4,1].PVAuto2 := 2400.0, [4,1].RangeMax := 100.0, [4,1].RampRate := 5.0, [4,1].RampRateSave := 5.0, [4,1].Deadband := 5.0, [4,1].RampTimer.PRE := 3600000, [4,1].StableTimer.PRE := 10000, [4,1].StableTime := 10, [4,1].PIDTimer.PRE := 250, [4,1].PIDTimer.ACC := 107, [4,1].PIDTimer.EN := 1, [4,1].PIDTimer.TT := 1, [4,1].CycleTimer.PRE := 2000, [4,1].PID.CTL := 67143552, [4,1].PID.SWM := 1, [4,1].PID.INI := 1, [4,1].PID.DVNA := 1, [4,1].PID.DVPA := 1, [4,1].PID.PVLA := 1, [4,1].PID.PVHA := 1, [4,1].PID.KP := 0.7, [4,1].PID.KI := 1.4, [4,1].PID.KD := 0.013, [4,1].PID.MAXS := 22.0, [4,1].PID.DB := 0.001, [4,1].PID.MAXO := 100.0, [4,1].PID.UPD := 0.25, [4,1].PID.MAXI := 22.0, [4,1].PID.MAXCV := 100.0, [4,1].PID.MAXTIE := 22.0, [4,1].PID.DATA[5] := 4.5454545, [4,1].PID.DATA[6] := 1.0, [4,1].PID.DATA[7] := 4.013, [4,1].PID.DATA[8] := 0.7, [4,1].PID.DATA[9] := 1.4, [4,1].PID.DATA[10] := 0.013, [4,1].PID.DATA[11] := 0.7, [4,1].PID.DATA[12] := 1.4, [4,1].PID.DATA[13] := 0.013, [4,1].PID.DATA[15] := 1.0, [4,1].PID.DATA[16] := 4.5454545, [4,1].KP[0] := 700.0, [4,1].KI[0] := 1400.0,
        [4,1].KD[0] := 13.0, [4,1].Auto1Cfg := 1, [4,1].Auto2Cfg := 1, [4,1].Auto1PVCfg := 10, [4,1].Auto2PVCfg := 42, [4,1].Auto1RangeMax := 22.0, [4,1].Auto2RangeMax := 9999.0, [4,2].Tag := 'FIC02', [4,2].Desc := 'Sec. Feed Pump Control', [4,2].LoopCfg := 1, [4,2].ManualEGU := '%', [4,2].Auto1EGU := 'LPM', [4,2].Auto2EGU := 'cm/h', [4,2].Interlock := 1, [4,2].Manual := 1, [4,2].DBOK := 1, [4,2].RampEnable := 1, [4,2].PIDEnable := 1, [4,2].ManualOSR := 1, [4,2].PVAuto2 := 2400.0, [4,2].RangeMax := 100.0, [4,2].RampRate := 5.0, [4,2].RampRateSave := 5.0, [4,2].RampStart := 75.0, [4,2].Deadband := 5.0, [4,2].RampTimer.PRE := 3600000, [4,2].StableTimer.PRE := 10000, [4,2].StableTime := 10, [4,2].PIDTimer.PRE := 250, [4,2].PIDTimer.ACC := 108, [4,2].PIDTimer.EN := 1, [4,2].PIDTimer.TT := 1, [4,2].CycleTimer.PRE := 2000, [4,2].PID.CTL := 67143552, [4,2].PID.SWM := 1, [4,2].PID.INI := 1, [4,2].PID.DVNA := 1, [4,2].PID.DVPA := 1, [4,2].PID.PVLA := 1, [4,2].PID.PVHA := 1, [4,2].PID.KP := 0.7, [4,2].PID.KI := 1.4, [4,2].PID.KD := 0.013, [4,2].PID.MAXS := 22.0, [4,2].PID.DB := 0.001, [4,2].PID.MAXO := 100.0, [4,2].PID.UPD := 0.25, [4,2].PID.MAXI := 22.0, [4,2].PID.MAXCV := 100.0, [4,2].PID.MAXTIE := 100.0, [4,2].PID.DATA[5] := 4.5454545, [4,2].PID.DATA[6] := 1.0, [4,2].PID.DATA[7] := 4.013, [4,2].PID.DATA[8] := 0.7, [4,2].PID.DATA[9] := 1.4, [4,2].PID.DATA[10] := 0.013, [4,2].PID.DATA[11] := 0.7, [4,2].PID.DATA[12] := 1.4, [4,2].PID.DATA[13] := 0.013, [4,2].PID.DATA[15] := 1.0,
        [4,2].PID.DATA[16] := 1.0, [4,2].KP[0] := 700.0, [4,2].KI[0] := 1400.0, [4,2].KD[0] := 13.0, [4,2].DisOSR := 1, [4,2].Auto1Cfg := 1, [4,2].Auto2Cfg := 1, [4,2].Auto1PVCfg := 12, [4,2].Auto2PVCfg := 43, [4,2].Auto1RangeMax := 22.0, [4,2].Auto2RangeMax := 9999.0, [4,2].OutputAddress := 1, [4,3].Tag := 'PCV12', [4,3].Desc := 'Post Column PCV012 Control', [4,3].LoopCfg := 1, [4,3].ManualEGU := '%', [4,3].Enable := 1, [4,3].Manual := 1, [4,3].Stable := 1, [4,3].DBOK := 1, [4,3].Status := 3, [4,3].RampEnable := 1, [4,3].PIDEnable := 1, [4,3].ManualOSR := 1, [4,3].RangeMax := 100.0, [4,3].RampRate := 5.0, [4,3].RampRateSave := 5.0, [4,3].RampStart := 98.0, [4,3].RampTimer.PRE := 3600000, [4,3].StableTimer.PRE := 2300, [4,3].StableTimer.ACC := 2354, [4,3].StableTimer.EN := 1, [4,3].StableTimer.DN := 1, [4,3].PIDTimer.PRE := 250, [4,3].PIDTimer.ACC := 108, [4,3].PIDTimer.EN := 1, [4,3].PIDTimer.TT := 1, [4,3].CycleTimer.PRE := 2000, [4,3].PID.CTL := 201361280, [4,3].PID.DOE := 1, [4,3].PID.SWM := 1, [4,3].PID.INI := 1, [4,3].PID.DVNA := 1, [4,3].PID.DVPA := 1, [4,3].PID.PVLA := 1, [4,3].PID.PVHA := 1, [4,3].PID.KP := 0.001, [4,3].PID.KI := 0.001, [4,3].PID.BIAS := 30.796, [4,3].PID.MAXS := 4095.0, [4,3].PID.MAXO := 100.0, [4,3].PID.UPD := 0.01, [4,3].PID.MAXI := 4095.0, [4,3].PID.MAXCV := 100.0, [4,3].PID.MAXTIE := 100.0, [4,3].PID.DATA[0] := -30.796, [4,3].PID.DATA[5] := 0.024420025, [4,3].PID.DATA[6] := 1.0, [4,3].PID.DATA[7] := 0.16, [4,3].PID.DATA[8] := 0.001,
        [4,3].PID.DATA[9] := 0.001, [4,3].PID.DATA[11] := 0.001, [4,3].PID.DATA[12] := 0.001, [4,3].PID.DATA[15] := 1.0, [4,3].PID.DATA[16] := 1.0, [4,3].OutputAddress := 2, [4,4].Tag := 'PCV10', [4,4].Desc := 'Line Pump1 PCV010 Control', [4,4].ManualEGU := '%', [4,4].Manual := 1, [4,4].Status := 3, [4,4].RampEnable := 1, [4,4].PIDEnable := 1, [4,4].RangeMax := 100.0, [4,4].RampRate := 0.5, [4,4].RampRateSave := 0.5, [4,4].RampStart := 3.443, [4,4].RampTimer.PRE := 3600000, [4,4].StableTimer.PRE := 5000, [4,4].PIDTimer.PRE := 250, [4,4].CycleTimer.PRE := 2000, [4,4].PID.CTL := 35652992, [4,4].PID.CA := 1, [4,4].PID.NOBC := 1, [4,4].PID.DVNA := 1, [4,4].PID.PVLA := 1, [4,4].PID.PVHA := 1, [4,4].PID.SP := 19.6, [4,4].PID.KP := 0.1, [4,4].PID.KI := 0.3, [4,4].PID.MAXS := 150.0, [4,4].PID.MAXO := 100.0, [4,4].PID.UPD := 0.25, [4,4].PID.ERR := -19.6, [4,4].PID.MAXI := 150.0, [4,4].PID.MAXCV := 100.0, [4,4].PID.MAXTIE := 100.0, [4,4].PID.DATA[0] := 1.3066667, [4,4].PID.DATA[3] := -19.6, [4,4].PID.DATA[4] := 19.6, [4,4].PID.DATA[5] := 0.6666667, [4,4].PID.DATA[6] := 1.0, [4,4].PID.DATA[7] := 4.0, [4,4].PID.DATA[8] := 0.1, [4,4].PID.DATA[9] := 0.3, [4,4].PID.DATA[11] := 0.1, [4,4].PID.DATA[12] := 0.3, [4,4].PID.DATA[15] := 1.0, [4,4].PID.DATA[16] := 1.0, [4,4].OutputAddress := 2, [4,5].Tag := 'PCV11', [4,5].Desc := 'Line Pump2 PCV011 Control', [4,5].ManualEGU := '%', [4,5].Manual := 1, [4,5].Status := 3, [4,5].RampEnable := 1, [4,5].PIDEnable := 1, [4,5].RangeMax := 100.0, [4,5].RampRate := 0.5, [4,5].RampRateSave := 0.5,
        [4,5].RampStart := 4.417, [4,5].RampTimer.PRE := 3600000, [4,5].StableTimer.PRE := 1500, [4,5].PIDTimer.PRE := 250, [4,5].CycleTimer.PRE := 2000, [4,5].PID.CTL := 134218624, [4,5].PID.DOE := 1, [4,5].PID.DVPA := 1, [4,5].PID.PVLA := 1, [4,5].PID.PVHA := 1, [4,5].PID.SP := 350.0, [4,5].PID.KP := 40.0, [4,5].PID.KI := 0.5, [4,5].PID.BIAS := -847.4798, [4,5].PID.MAXS := 550.0, [4,5].PID.MAXO := 100.0, [4,5].PID.UPD := 0.25, [4,5].PID.ERR := 350.0, [4,5].PID.MAXI := 550.0, [4,5].PID.MAXCV := 100.0, [4,5].PID.MAXTIE := 100.0, [4,5].PID.DATA[0] := -1697.9749, [4,5].PID.DATA[1] := 1018.1818, [4,5].PID.DATA[3] := 350.0, [4,5].PID.DATA[4] := 350.0, [4,5].PID.DATA[5] := 0.18181819, [4,5].PID.DATA[6] := 1.0, [4,5].PID.DATA[7] := 4.0, [4,5].PID.DATA[8] := 40.0, [4,5].PID.DATA[9] := 0.5, [4,5].PID.DATA[11] := 40.0, [4,5].PID.DATA[12] := 0.5, [4,5].PID.DATA[15] := 1.0, [4,5].PID.DATA[16] := 1.0, [4,5].OutputAddress := 3, [4,6].StableTimer.PRE := 15000, [4,6].PIDTimer.EN := 1, [4,6].PIDTimer.TT := 1, [4,6].CycleTimer.PRE := 5000, [4,6].PID.CTL := 16810624, [4,6].PID.MO := 1, [4,6].PID.INI := 1, [4,6].PID.DVPA := 1, [4,6].PID.PVHA := 1, [4,6].PID.SP := 10.0, [4,6].PID.KP := 0.3, [4,6].PID.KI := 0.3, [4,6].PID.MAXS := 200.0, [4,6].PID.SO := 3.074094, [4,6].PID.MAXO := 100.0, [4,6].PID.UPD := 0.25, [4,6].PID.PV := 1.488363, [4,6].PID.ERR := 8.511638, [4,6].PID.OUT := 3.074094, [4,6].PID.MAXI := 200.0, [4,6].PID.TIE := 3.074094, [4,6].PID.MAXCV := 200.0, [4,6].PID.MAXTIE := 200.0, [4,6].PID.DATA[0] := 1.797348, [4,6].PID.DATA[1] := -11.9069,
        [4,6].PID.DATA[2] := 1.488363, [4,6].PID.DATA[3] := 8.511638, [4,6].PID.DATA[4] := 10.0, [4,6].PID.DATA[5] := 0.5, [4,6].PID.DATA[6] := 1.0, [4,6].PID.DATA[7] := 4.0, [4,6].PID.DATA[8] := 0.3, [4,6].PID.DATA[9] := 0.3, [4,6].PID.DATA[11] := 0.3, [4,6].PID.DATA[12] := 0.3, [4,6].PID.DATA[15] := 2.0, [4,6].PID.DATA[16] := 0.5, [4,7].StableTimer.PRE := 200, [4,7].PIDTimer.PRE := 250, [4,7].PIDTimer.EN := 1, [4,7].PIDTimer.TT := 1, [4,7].CycleTimer.PRE := 10000, [4,7].PID.CTL := 16810880, [4,7].PID.MO := 1, [4,7].PID.INI := 1, [4,7].PID.DVPA := 1, [4,7].PID.PVLA := 1, [4,7].PID.PVHA := 1, [4,7].PID.SP := 10.0, [4,7].PID.KP := 2.0, [4,7].PID.KI := 0.2, [4,7].PID.KD := 0.3, [4,7].PID.BIAS := 50.0, [4,7].PID.DB := 0.01, [4,7].PID.SO := 80.0, [4,7].PID.MAXO := 100.0, [4,7].PID.UPD := 0.25, [4,7].PID.ERR := 10.0, [4,7].PID.OUT := 80.0, [4,7].PID.TIE := 80.0, [4,7].PID.MAXCV := 100.0, [4,7].PID.MAXTIE := 100.0, [4,7].PID.DATA[0] := 29.511597, [4,7].PID.DATA[3] := 10.0, [4,7].PID.DATA[4] := 10.0, [4,7].PID.DATA[5] := 0.024420025, [4,7].PID.DATA[6] := 1.0, [4,7].PID.DATA[7] := 4.3, [4,7].PID.DATA[8] := 2.0, [4,7].PID.DATA[9] := 0.2, [4,7].PID.DATA[10] := 0.3, [4,7].PID.DATA[11] := 2.0, [4,7].PID.DATA[12] := 0.2, [4,7].PID.DATA[13] := 0.3, [4,7].PID.DATA[15] := 1.0, [4,7].PID.DATA[16] := 1.0, [4,8].StableTimer.PRE := 15000, [4,8].PIDTimer.PRE := 250, [4,8].CycleTimer.PRE := 20000, [4,8].PID.CTL := 33555584, [4,8].PID.CA := 1, [4,8].PID.DVNA := 1, [4,8].PID.PVHA := 1, [4,8].PID.SP := 27.0, [4,8].PID.KP := 1.0,
        [4,8].PID.KI := 0.1, [4,8].PID.MAXS := 100.0, [4,8].PID.MAXO := 100.0, [4,8].PID.UPD := 0.25, [4,8].PID.PV := 18.2328, [4,8].PID.ERR := -8.767202, [4,8].PID.MAXI := 100.0, [4,8].PID.MAXCV := 100.0, [4,8].PID.MAXTIE := 100.0, [4,8].PID.DATA[0] := 8.767202, [4,8].PID.DATA[1] := 291.7248, [4,8].PID.DATA[2] := 18.2328, [4,8].PID.DATA[3] := -8.767202, [4,8].PID.DATA[4] := 27.0, [4,8].PID.DATA[5] := 1.0, [4,8].PID.DATA[6] := 1.0, [4,8].PID.DATA[7] := 4.0, [4,8].PID.DATA[8] := 1.0, [4,8].PID.DATA[9] := 0.1, [4,8].PID.DATA[11] := 1.0, [4,8].PID.DATA[12] := 0.1, [4,8].PID.DATA[15] := 1.0, [4,8].PID.DATA[16] := 1.0, [4,11].RampTimer.PRE := 100000, [4,11].StableTimer.PRE := 200, [4,11].PIDTimer.PRE := 250, [4,11].PIDTimer.ACC := 230, [4,11].PIDTimer.EN := 1, [4,11].PIDTimer.TT := 1, [4,11].PID.CTL := 67142528, [4,11].PID.SWM := 1, [4,11].PID.INI := 1, [4,11].PID.DVPA := 1, [4,11].PID.PVLA := 1, [4,11].PID.PVHA := 1, [4,11].PID.SP := 0.20000005, [4,11].PID.KP := 0.1, [4,11].PID.KI := 0.1, [4,11].PID.BIAS := 23.09767, [4,11].PID.DB := 0.001, [4,11].PID.MAXO := 100.0, [4,11].PID.UPD := 0.25, [4,11].PID.ERR := 0.20000005, [4,11].PID.MAXCV := 100.0, [4,11].PID.MAXTIE := 100.0, [4,11].PID.DATA[0] := -23.098158, [4,11].PID.DATA[3] := 0.20000005, [4,11].PID.DATA[4] := 0.20000005, [4,11].PID.DATA[5] := 0.024420025, [4,11].PID.DATA[6] := 1.0, [4,11].PID.DATA[7] := 4.0, [4,11].PID.DATA[8] := 0.1, [4,11].PID.DATA[9] := 0.1, [4,11].PID.DATA[11] := 0.1, [4,11].PID.DATA[12] := 0.1, [4,11].PID.DATA[15] := 1.0, [4,11].PID.DATA[16] := 1.0, [4,13].RampTimer.PRE := 3600000, [4,13].StableTimer.PRE := 2000, [4,13].PIDTimer.PRE := 10000,
        [4,13].PIDTimer.EN := 1, [4,13].PIDTimer.TT := 1, [4,13].PID.CTL := 305173120, [4,13].PID.PVT := 1, [4,13].PID.CA := 1, [4,13].PID.NOBC := 1, [4,13].PID.NOZC := 1, [4,13].PID.INI := 1, [4,13].PID.OLH := 1, [4,13].PID.DVPA := 1, [4,13].PID.PVHA := 1, [4,13].PID.KP := 0.2, [4,13].PID.KI := 0.08, [4,13].PID.MAXS := 100.0, [4,13].PID.DB := 1.0, [4,13].PID.SO := 100.0, [4,13].PID.MAXO := 100.0, [4,13].PID.UPD := 0.01, [4,13].PID.PV := 43.925232, [4,13].PID.ERR := 43.925232, [4,13].PID.OUT := 100.0, [4,13].PID.MAXI := 100.0, [4,13].PID.TIE := 2.4420025, [4,13].PID.MAXCV := 100.0, [4,13].PID.MAXTIE := 4095.0, [4,13].PID.DATA[0] := 100.0, [4,13].PID.DATA[1] := 702.8037, [4,13].PID.DATA[2] := 43.925232, [4,13].PID.DATA[3] := 43.925232, [4,13].PID.DATA[5] := 1.0, [4,13].PID.DATA[6] := 1.0, [4,13].PID.DATA[7] := 0.16, [4,13].PID.DATA[8] := 0.2, [4,13].PID.DATA[9] := 0.08, [4,13].PID.DATA[11] := 0.2, [4,13].PID.DATA[12] := 0.08, [4,13].PID.DATA[15] := 1.0, [4,13].PID.DATA[16] := 0.024420025, [5,0].RampTimer.PRE := 3600000, [5,0].StableTimer.PRE := 5000, [5,0].PIDTimer.PRE := 250, [5,0].PIDTimer.ACC := 100, [5,0].PIDTimer.EN := 1, [5,0].PIDTimer.TT := 1, [5,0].PID.CTL := 25199488, [5,0].PID.MO := 1, [5,0].PID.PE := 1, [5,0].PID.INI := 1, [5,0].PID.DVPA := 1, [5,0].PID.PVLA := 1, [5,0].PID.PVHA := 1, [5,0].PID.SP := 66.66666, [5,0].PID.KP := 0.5, [5,0].PID.KI := 0.1, [5,0].PID.MAXS := 200.0, [5,0].PID.SO := 10.0, [5,0].PID.MAXO := 100.0, [5,0].PID.MINO := 10.0, [5,0].PID.UPD := 0.25, [5,0].PID.ERR := 66.66666,
        [5,0].PID.OUT := 10.0, [5,0].PID.MAXI := 200.0, [5,0].PID.TIE := 10.0, [5,0].PID.MAXCV := 100.0, [5,0].PID.MAXTIE := 100.0, [5,0].PID.DATA[0] := -6.666666, [5,0].PID.DATA[3] := 66.66666, [5,0].PID.DATA[4] := 66.66666, [5,0].PID.DATA[5] := 0.5, [5,0].PID.DATA[6] := 1.0, [5,0].PID.DATA[7] := 4.0, [5,0].PID.DATA[8] := 0.5, [5,0].PID.DATA[9] := 0.1, [5,0].PID.DATA[11] := 0.5, [5,0].PID.DATA[12] := 0.08333334, [5,0].PID.DATA[15] := 1.0, [5,0].PID.DATA[16] := 1.0, [5,1].Tag := 'FIC01', [5,1].Desc := 'Prim. Feed Pump Control', [5,1].LoopCfg := 1, [5,1].ManualEGU := '%', [5,1].Auto1EGU := 'LPM', [5,1].Auto2EGU := 'cm/h', [5,1].Manual := 1, [5,1].DBOK := 1, [5,1].RampEnable := 1, [5,1].PIDEnable := 1, [5,1].ManualOSR := 1, [5,1].PVAuto2 := 2400.0, [5,1].RangeMax := 100.0, [5,1].RampRate := 5.0, [5,1].RampRateSave := 5.0, [5,1].Deadband := 5.0, [5,1].RampTimer.PRE := 3600000, [5,1].StableTimer.PRE := 10000, [5,1].StableTime := 10, [5,1].PIDTimer.PRE := 250, [5,1].PIDTimer.EN := 1, [5,1].PIDTimer.TT := 1, [5,1].CycleTimer.PRE := 2000, [5,1].PID.CTL := 67143552, [5,1].PID.SWM := 1, [5,1].PID.INI := 1, [5,1].PID.DVNA := 1, [5,1].PID.DVPA := 1, [5,1].PID.PVLA := 1, [5,1].PID.PVHA := 1, [5,1].PID.KP := 0.7, [5,1].PID.KI := 1.4, [5,1].PID.KD := 0.013, [5,1].PID.DB := 0.001, [5,1].PID.MAXO := 100.0, [5,1].PID.UPD := 0.25, [5,1].PID.MAXCV := 100.0, [5,1].PID.DATA[5] := 0.024420025, [5,1].PID.DATA[6] := 1.0, [5,1].PID.DATA[7] := 4.013, [5,1].PID.DATA[8] := 0.7, [5,1].PID.DATA[9] := 1.4, [5,1].PID.DATA[10] := 0.013,
        [5,1].PID.DATA[11] := 0.7, [5,1].PID.DATA[12] := 1.4, [5,1].PID.DATA[13] := 0.013, [5,1].PID.DATA[15] := 1.0, [5,1].PID.DATA[16] := 1.0, [5,1].KP[0] := 700.0, [5,1].KI[0] := 1400.0, [5,1].KD[0] := 13.0, [5,1].Auto1Cfg := 1, [5,1].Auto2Cfg := 1, [5,1].Auto1PVCfg := 10, [5,1].Auto2PVCfg := 42, [5,1].Auto2RangeMax := 5.0, [5,2].Tag := 'FIC02', [5,2].Desc := 'Sec. Feed Pump Control', [5,2].LoopCfg := 1, [5,2].ManualEGU := '%', [5,2].Auto1EGU := 'LPM', [5,2].Auto2EGU := 'cm/h', [5,2].Interlock := 1, [5,2].Manual := 1, [5,2].DBOK := 1, [5,2].RampEnable := 1, [5,2].PIDEnable := 1, [5,2].ManualOSR := 1, [5,2].PVAuto2 := 2400.0, [5,2].RangeMax := 100.0, [5,2].RampRate := 5.0, [5,2].RampRateSave := 5.0, [5,2].RampStart := 75.0, [5,2].Deadband := 5.0, [5,2].RampTimer.PRE := 3600000, [5,2].StableTimer.PRE := 10000, [5,2].StableTime := 10, [5,2].PIDTimer.PRE := 250, [5,2].PIDTimer.EN := 1, [5,2].PIDTimer.TT := 1, [5,2].CycleTimer.PRE := 2000, [5,2].PID.CTL := 67143552, [5,2].PID.SWM := 1, [5,2].PID.INI := 1, [5,2].PID.DVNA := 1, [5,2].PID.DVPA := 1, [5,2].PID.PVLA := 1, [5,2].PID.PVHA := 1, [5,2].PID.KP := 0.7, [5,2].PID.KI := 1.4, [5,2].PID.KD := 0.013, [5,2].PID.MAXS := 50.0, [5,2].PID.DB := 0.001, [5,2].PID.MAXO := 100.0, [5,2].PID.UPD := 0.25, [5,2].PID.MAXI := 50.0, [5,2].PID.MAXCV := 100.0, [5,2].PID.MAXTIE := 100.0, [5,2].PID.DATA[5] := 2.0, [5,2].PID.DATA[6] := 1.0, [5,2].PID.DATA[7] := 4.013, [5,2].PID.DATA[8] := 0.7, [5,2].PID.DATA[9] := 1.4,
        [5,2].PID.DATA[10] := 0.013, [5,2].PID.DATA[11] := 0.7, [5,2].PID.DATA[12] := 1.4, [5,2].PID.DATA[13] := 0.013, [5,2].PID.DATA[15] := 1.0, [5,2].PID.DATA[16] := 1.0, [5,2].KP[0] := 700.0, [5,2].KI[0] := 1400.0, [5,2].KD[0] := 13.0, [5,2].DisOSR := 1, [5,2].Auto1Cfg := 1, [5,2].Auto2Cfg := 1, [5,2].Auto1PVCfg := 12, [5,2].Auto2PVCfg := 43, [5,2].Auto1RangeMax := 50.0, [5,2].Auto2RangeMax := 99999.0, [5,2].OutputAddress := 1, [5,3].Tag := 'PCV12', [5,3].Desc := 'Post Column PCV012 Control', [5,3].LoopCfg := 1, [5,3].ManualEGU := '%', [5,3].Enable := 1, [5,3].Manual := 1, [5,3].Stable := 1, [5,3].DBOK := 1, [5,3].Status := 3, [5,3].RampEnable := 1, [5,3].PIDEnable := 1, [5,3].ManualOSR := 1, [5,3].RangeMax := 100.0, [5,3].RampRate := 5.0, [5,3].RampRateSave := 5.0, [5,3].RampStart := 98.0, [5,3].RampTimer.PRE := 3600000, [5,3].StableTimer.PRE := 2300, [5,3].StableTimer.ACC := 2354, [5,3].StableTimer.EN := 1, [5,3].StableTimer.DN := 1, [5,3].PIDTimer.PRE := 250, [5,3].PIDTimer.EN := 1, [5,3].PIDTimer.TT := 1, [5,3].CycleTimer.PRE := 2000, [5,3].PID.CTL := 201361280, [5,3].PID.DOE := 1, [5,3].PID.SWM := 1, [5,3].PID.INI := 1, [5,3].PID.DVNA := 1, [5,3].PID.DVPA := 1, [5,3].PID.PVLA := 1, [5,3].PID.PVHA := 1, [5,3].PID.KP := 0.001, [5,3].PID.KI := 0.001, [5,3].PID.BIAS := 30.796, [5,3].PID.MAXS := 4095.0, [5,3].PID.MAXO := 100.0, [5,3].PID.UPD := 0.01, [5,3].PID.MAXI := 4095.0, [5,3].PID.MAXCV := 100.0, [5,3].PID.MAXTIE := 100.0, [5,3].PID.DATA[0] := -30.796,
        [5,3].PID.DATA[5] := 0.024420025, [5,3].PID.DATA[6] := 1.0, [5,3].PID.DATA[7] := 0.16, [5,3].PID.DATA[8] := 0.001, [5,3].PID.DATA[9] := 0.001, [5,3].PID.DATA[11] := 0.001, [5,3].PID.DATA[12] := 0.001, [5,3].PID.DATA[15] := 1.0, [5,3].PID.DATA[16] := 1.0, [5,3].OutputAddress := 2, [5,4].Tag := 'PCV10', [5,4].Desc := 'Line Pump1 PCV010 Control', [5,4].ManualEGU := '%', [5,4].Manual := 1, [5,4].Status := 3, [5,4].RampEnable := 1, [5,4].PIDEnable := 1, [5,4].RangeMax := 100.0, [5,4].RampRate := 0.5, [5,4].RampRateSave := 0.5, [5,4].RampStart := 3.443, [5,4].RampTimer.PRE := 3600000, [5,4].StableTimer.PRE := 5000, [5,4].PIDTimer.PRE := 250, [5,4].CycleTimer.PRE := 2000, [5,4].PID.CTL := 35652992, [5,4].PID.CA := 1, [5,4].PID.NOBC := 1, [5,4].PID.DVNA := 1, [5,4].PID.PVLA := 1, [5,4].PID.PVHA := 1, [5,4].PID.SP := 19.6, [5,4].PID.KP := 0.1, [5,4].PID.KI := 0.3, [5,4].PID.MAXS := 150.0, [5,4].PID.MAXO := 100.0, [5,4].PID.UPD := 0.25, [5,4].PID.ERR := -19.6, [5,4].PID.MAXI := 150.0, [5,4].PID.MAXCV := 100.0, [5,4].PID.MAXTIE := 100.0, [5,4].PID.DATA[0] := 1.3066667, [5,4].PID.DATA[3] := -19.6, [5,4].PID.DATA[4] := 19.6, [5,4].PID.DATA[5] := 0.6666667, [5,4].PID.DATA[6] := 1.0, [5,4].PID.DATA[7] := 4.0, [5,4].PID.DATA[8] := 0.1, [5,4].PID.DATA[9] := 0.3, [5,4].PID.DATA[11] := 0.1, [5,4].PID.DATA[12] := 0.3, [5,4].PID.DATA[15] := 1.0, [5,4].PID.DATA[16] := 1.0, [5,4].OutputAddress := 2, [5,5].Tag := 'PCV11', [5,5].Desc := 'Line Pump2 PCV011 Control', [5,5].ManualEGU := '%', [5,5].Manual := 1, [5,5].Status := 3, [5,5].RampEnable := 1,
        [5,5].PIDEnable := 1, [5,5].RangeMax := 100.0, [5,5].RampRate := 0.5, [5,5].RampRateSave := 0.5, [5,5].RampStart := 4.417, [5,5].RampTimer.PRE := 3600000, [5,5].StableTimer.PRE := 1500, [5,5].PIDTimer.PRE := 250, [5,5].CycleTimer.PRE := 2000, [5,5].PID.CTL := 134218624, [5,5].PID.DOE := 1, [5,5].PID.DVPA := 1, [5,5].PID.PVLA := 1, [5,5].PID.PVHA := 1, [5,5].PID.SP := 350.0, [5,5].PID.KP := 40.0, [5,5].PID.KI := 0.5, [5,5].PID.BIAS := -847.4798, [5,5].PID.MAXS := 550.0, [5,5].PID.MAXO := 100.0, [5,5].PID.UPD := 0.25, [5,5].PID.ERR := 350.0, [5,5].PID.MAXI := 550.0, [5,5].PID.MAXCV := 100.0, [5,5].PID.MAXTIE := 100.0, [5,5].PID.DATA[0] := -1697.9749, [5,5].PID.DATA[1] := 1018.1818, [5,5].PID.DATA[3] := 350.0, [5,5].PID.DATA[4] := 350.0, [5,5].PID.DATA[5] := 0.18181819, [5,5].PID.DATA[6] := 1.0, [5,5].PID.DATA[7] := 4.0, [5,5].PID.DATA[8] := 40.0, [5,5].PID.DATA[9] := 0.5, [5,5].PID.DATA[11] := 40.0, [5,5].PID.DATA[12] := 0.5, [5,5].PID.DATA[15] := 1.0, [5,5].PID.DATA[16] := 1.0, [5,5].OutputAddress := 3, [5,6].StableTimer.PRE := 15000, [5,6].PIDTimer.EN := 1, [5,6].PIDTimer.TT := 1, [5,6].CycleTimer.PRE := 5000, [5,6].PID.CTL := 16810624, [5,6].PID.MO := 1, [5,6].PID.INI := 1, [5,6].PID.DVPA := 1, [5,6].PID.PVHA := 1, [5,6].PID.SP := 10.0, [5,6].PID.KP := 0.3, [5,6].PID.KI := 0.3, [5,6].PID.MAXS := 200.0, [5,6].PID.SO := 3.074094, [5,6].PID.MAXO := 100.0, [5,6].PID.UPD := 0.25, [5,6].PID.PV := 1.488363, [5,6].PID.ERR := 8.511638, [5,6].PID.OUT := 3.074094, [5,6].PID.MAXI := 200.0, [5,6].PID.TIE := 3.074094,
        [5,6].PID.MAXCV := 200.0, [5,6].PID.MAXTIE := 200.0, [5,6].PID.DATA[0] := 1.797348, [5,6].PID.DATA[1] := -11.9069, [5,6].PID.DATA[2] := 1.488363, [5,6].PID.DATA[3] := 8.511638, [5,6].PID.DATA[4] := 10.0, [5,6].PID.DATA[5] := 0.5, [5,6].PID.DATA[6] := 1.0, [5,6].PID.DATA[7] := 4.0, [5,6].PID.DATA[8] := 0.3, [5,6].PID.DATA[9] := 0.3, [5,6].PID.DATA[11] := 0.3, [5,6].PID.DATA[12] := 0.3, [5,6].PID.DATA[15] := 2.0, [5,6].PID.DATA[16] := 0.5, [5,7].StableTimer.PRE := 200, [5,7].PIDTimer.PRE := 250, [5,7].PIDTimer.EN := 1, [5,7].PIDTimer.TT := 1, [5,7].CycleTimer.PRE := 10000, [5,7].PID.CTL := 16810880, [5,7].PID.MO := 1, [5,7].PID.INI := 1, [5,7].PID.DVPA := 1, [5,7].PID.PVLA := 1, [5,7].PID.PVHA := 1, [5,7].PID.SP := 10.0, [5,7].PID.KP := 2.0, [5,7].PID.KI := 0.2, [5,7].PID.KD := 0.3, [5,7].PID.BIAS := 50.0, [5,7].PID.DB := 0.01, [5,7].PID.SO := 80.0, [5,7].PID.MAXO := 100.0, [5,7].PID.UPD := 0.25, [5,7].PID.ERR := 10.0, [5,7].PID.OUT := 80.0, [5,7].PID.TIE := 80.0, [5,7].PID.MAXCV := 100.0, [5,7].PID.MAXTIE := 100.0, [5,7].PID.DATA[0] := 29.511597, [5,7].PID.DATA[3] := 10.0, [5,7].PID.DATA[4] := 10.0, [5,7].PID.DATA[5] := 0.024420025, [5,7].PID.DATA[6] := 1.0, [5,7].PID.DATA[7] := 4.3, [5,7].PID.DATA[8] := 2.0, [5,7].PID.DATA[9] := 0.2, [5,7].PID.DATA[10] := 0.3, [5,7].PID.DATA[11] := 2.0, [5,7].PID.DATA[12] := 0.2, [5,7].PID.DATA[13] := 0.3, [5,7].PID.DATA[15] := 1.0, [5,7].PID.DATA[16] := 1.0, [5,8].StableTimer.PRE := 15000, [5,8].PIDTimer.PRE := 250, [5,8].CycleTimer.PRE := 20000, [5,8].PID.CTL := 33555584, [5,8].PID.CA := 1,
        [5,8].PID.DVNA := 1, [5,8].PID.PVHA := 1, [5,8].PID.SP := 27.0, [5,8].PID.KP := 1.0, [5,8].PID.KI := 0.1, [5,8].PID.MAXS := 100.0, [5,8].PID.MAXO := 100.0, [5,8].PID.UPD := 0.25, [5,8].PID.PV := 18.2328, [5,8].PID.ERR := -8.767202, [5,8].PID.MAXI := 100.0, [5,8].PID.MAXCV := 100.0, [5,8].PID.MAXTIE := 100.0, [5,8].PID.DATA[0] := 8.767202, [5,8].PID.DATA[1] := 291.7248, [5,8].PID.DATA[2] := 18.2328, [5,8].PID.DATA[3] := -8.767202, [5,8].PID.DATA[4] := 27.0, [5,8].PID.DATA[5] := 1.0, [5,8].PID.DATA[6] := 1.0, [5,8].PID.DATA[7] := 4.0, [5,8].PID.DATA[8] := 1.0, [5,8].PID.DATA[9] := 0.1, [5,8].PID.DATA[11] := 1.0, [5,8].PID.DATA[12] := 0.1, [5,8].PID.DATA[15] := 1.0, [5,8].PID.DATA[16] := 1.0, [5,11].RampTimer.PRE := 100000, [5,11].StableTimer.PRE := 200, [5,11].PIDTimer.PRE := 250, [5,11].PIDTimer.ACC := 230, [5,11].PIDTimer.EN := 1, [5,11].PIDTimer.TT := 1, [5,11].PID.CTL := 67142528, [5,11].PID.SWM := 1, [5,11].PID.INI := 1, [5,11].PID.DVPA := 1, [5,11].PID.PVLA := 1, [5,11].PID.PVHA := 1, [5,11].PID.SP := 0.20000005, [5,11].PID.KP := 0.1, [5,11].PID.KI := 0.1, [5,11].PID.BIAS := 23.09767, [5,11].PID.DB := 0.001, [5,11].PID.MAXO := 100.0, [5,11].PID.UPD := 0.25, [5,11].PID.ERR := 0.20000005, [5,11].PID.MAXCV := 100.0, [5,11].PID.MAXTIE := 100.0, [5,11].PID.DATA[0] := -23.098158, [5,11].PID.DATA[3] := 0.20000005, [5,11].PID.DATA[4] := 0.20000005, [5,11].PID.DATA[5] := 0.024420025, [5,11].PID.DATA[6] := 1.0, [5,11].PID.DATA[7] := 4.0, [5,11].PID.DATA[8] := 0.1, [5,11].PID.DATA[9] := 0.1, [5,11].PID.DATA[11] := 0.1, [5,11].PID.DATA[12] := 0.1, [5,11].PID.DATA[15] := 1.0,
        [5,11].PID.DATA[16] := 1.0, [5,13].RampTimer.PRE := 3600000, [5,13].StableTimer.PRE := 2000, [5,13].PIDTimer.PRE := 10000, [5,13].PIDTimer.EN := 1, [5,13].PIDTimer.TT := 1, [5,13].PID.CTL := 305173120, [5,13].PID.PVT := 1, [5,13].PID.CA := 1, [5,13].PID.NOBC := 1, [5,13].PID.NOZC := 1, [5,13].PID.INI := 1, [5,13].PID.OLH := 1, [5,13].PID.DVPA := 1, [5,13].PID.PVHA := 1, [5,13].PID.KP := 0.2, [5,13].PID.KI := 0.08, [5,13].PID.MAXS := 100.0, [5,13].PID.DB := 1.0, [5,13].PID.SO := 100.0, [5,13].PID.MAXO := 100.0, [5,13].PID.UPD := 0.01, [5,13].PID.PV := 43.925232, [5,13].PID.ERR := 43.925232, [5,13].PID.OUT := 100.0, [5,13].PID.MAXI := 100.0, [5,13].PID.TIE := 2.4420025, [5,13].PID.MAXCV := 100.0, [5,13].PID.MAXTIE := 4095.0, [5,13].PID.DATA[0] := 100.0, [5,13].PID.DATA[1] := 702.8037, [5,13].PID.DATA[2] := 43.925232, [5,13].PID.DATA[3] := 43.925232, [5,13].PID.DATA[5] := 1.0, [5,13].PID.DATA[6] := 1.0, [5,13].PID.DATA[7] := 0.16, [5,13].PID.DATA[8] := 0.2, [5,13].PID.DATA[9] := 0.08, [5,13].PID.DATA[11] := 0.2, [5,13].PID.DATA[12] := 0.08, [5,13].PID.DATA[15] := 1.0, [5,13].PID.DATA[16] := 0.024420025);
   ControlLoop_TIC101 : ALIAS FOR ControlLoop[7];
   ControlLoop_TIC101Alarm : ALIAS FOR AlarmDeviation[7];
   CPU_Scanning : BOOL := 1;   // System Scanning Flag
   CriteriaFlag : CriteriaFlag;   // Criteria Flag used in CCP Recipe
   DerivedData : DerivedData := (HOLDUP := 6.128, FI101Q := 100.0, FI201Q := 100.0, FI401Q := 100.0, FI101K := 1.0, FI201K := 1.0, FI401K := 1.0);   // Derived data (user input and calculated values)
   DF24VDC : ALIAS FOR DigitalPoint[4];
   DF24VDCPC : ALIAS FOR DigitalPoint[25];
   DF3PHP003 : ALIAS FOR DigitalPoint[27];
   DF48MIX : ALIAS FOR DigitalPoint[26];
   DF48P001 : ALIAS FOR DigitalPoint[23];
   DF48P002 : ALIAS FOR DigitalPoint[24];
   DI1 : ALIAS FOR DigitalPoint[34];
   DI2 : ALIAS FOR DigitalPoint[35];
   DI3 : ALIAS FOR DigitalPoint[36];
   DI4 : ALIAS FOR DigitalPoint[37];
   DI5 : ALIAS FOR DigitalPoint[38];
   DI6 : ALIAS FOR DigitalPoint[39];
   DI7 : ALIAS FOR DigitalPoint[40];
   DI8 : ALIAS FOR DigitalPoint[41];
   Diafiltration : Diafiltration := (Diaf_Init := 161.77638, Diaf_Final_Volume := 10.2, LogDiafTimer.PRE := 3000);
   DigitalInput : BOOL[256] := ([5] := 1, [6] := 1, [7] := 1, [8] := 1, [9] := 1, [10] := 1, [21] := 1, [22] := 1, [100] := 1, [104] := 1, [106] := 1, [111] := 1, [131] := 1);   // Digital Input Array these bits are copied from Input cards.
   DigitalOutput : BOOL[256] := ([1] := 1, [2] := 1, [5] := 1, [6] := 1, [11] := 1, [12] := 1, [14] := 1, [180] := 1, [181] := 1);   // Digital Output Array these bits are sent to output cards.
        [13]   // Disconnect multicontact
        [14]   // Powerup C8000
        [7]   // UV Auto Zero
        [17]   // Mixer Alarm Reset
        [18]   // Feed Tank Tare
        [10]   // Unlock CS
        [11]   // Lock CS
        [12]   // Connect multicontact
        [21]   // Tare Feed Pump Pressure
        [8]   // Start pump P001
        [15]   // Start pump P003
        [16]   // Start Mixer MIX101
        [19]   // Feed Tank Clear Tare
        [1]   // System powered-up
        [20]   // Bath TCU Enable
        [22]   // Tare Retentate Pressure
        [26]   // Tare Feed Tank Pressure
        [23]   // Tare Filtrate Pressure
        [24]   // Tare Transfer Pump Pressure
        [25]   // Inflate Bag
        [5]   // Lighting banner red Smart
        [27]   // Weight Zero
        [2]   // BUZZER
        [32]   // Valve XV001
        [33]   // Valve XV002
        [34]   // Valve XV003
        [35]   // Valve XV004
        [36]   // Valve XV005
        [37]   // Valve XV006
        [38]   // Valve XV007
        [39]   // Valve XV101
        [3]   // Lighting banner green Smart
        [40]   // Valve XV102
        [41]   // Valve XV401
        [42]   // Valve XV402
        [43]   // Valve XV403
        [44]   // Valve XV404
        [45]   // Valve XV405
        [46]   // Valve XV406
        [47]   // Valve XV201
        [48]   // Valve XV202
        [49]   // Valve XV701
        [4]   // Lighting banner green Pcart
        [50]   // Valve XV702
        [51]   // Valve XV703
        [52]   // Valve XV704
        [6]   // Lighting banner red Pcart
        [80]   // DO1
        [81]   // DO2
        [82]   // DO3
        [83]   // DO4
        [84]   // DO5
        [85]   // DO6
        [86]   // DO7
        [87]   // DO8
        [9]   // Start pump P002
        [0]   // Re-established system
   DigitalPoint : DigitalPoint[150] := ([0].Tag := 'PSL602', [0].AlarmCurrentValue := 1, [0].Override := 1, [0].DelayTimer.PRE := 5000, [0].DelayTimer.ACC := 5040, [0].DelayTimer.EN := 1, [0].DelayTimer.DN := 1, [0].DelayTimerSP := 5, [0].Priority := 1, [0].EnableCfg := 1, [0].ActiveStateCFg := 1, [0].RealInputCfg := 1, [0].AlarmCfg := 1, [0].OverrideCfg := 1, [0].PriorityCfg := 1, [1].Tag := 'XS001', [1].AlarmCurrentValue := 1, [1].Override := 1, [1].Condition2 := 1, [1].DelayTimer.PRE := 5000, [1].DelayTimer.ACC := 5041, [1].DelayTimer.EN := 1, [1].DelayTimer.DN := 1, [1].DelayTimerSP := 5, [1].Priority := 1, [1].EnableCfg := 1, [1].ActiveStateCFg := 1, [1].RealInputCfg := 1, [1].InputAddressCfg := 1, [1].AlarmCfg := 1, [1].OverrideCfg := 1, [1].PriorityCfg := 1, [2].Tag := 'XS006', [2].AlarmCurrentValue := 1, [2].Alarm := 1, [2].Mimic := 4, [2].DelayTimer.ACC := 51, [2].DelayTimer.EN := 1, [2].DelayTimer.DN := 1, [2].Priority := 1, [2].EnableCfg := 1, [2].ActiveStateCFg := 1, [2].RealInputCfg := 1, [2].InputAddressCfg := 2, [2].AlarmCfg := 1, [2].AlarmONS := 1, [3].Tag := 'ES001', [3].DelayTimer.PRE := 2000, [3].DelayTimerSP := 2, [3].EnableCfg := 1, [3].ActiveStateCFg := 1, [3].RealInputCfg := 1, [3].InputAddressCfg := 3, [4].Tag := 'PSH001', [4].AlarmCurrentValue := 1, [4].Override := 1, [4].DelayTimer.PRE := 1000, [4].DelayTimer.ACC := 1030, [4].DelayTimer.EN := 1, [4].DelayTimer.DN := 1,
        [4].DelayTimerSP := 1, [4].Priority := 1, [4].EnableCfg := 1, [4].ActiveStateCFg := 1, [4].RealInputCfg := 1, [4].InputAddressCfg := 4, [4].AlarmCfg := 1, [4].OverrideCfg := 1, [4].PriorityCfg := 1, [5].Tag := 'PSH401', [5].CurrentValue := 1, [5].Override := 1, [5].Mimic := 1, [5].DelayTimer.PRE := 1000, [5].DelayTimerSP := 1, [5].Priority := 1, [5].EnableCfg := 1, [5].ActiveStateCFg := 1, [5].RealInputCfg := 1, [5].InputAddressCfg := 5, [5].AlarmCfg := 1, [5].OverrideCfg := 1, [5].PriorityCfg := 1, [6].Tag := 'XS002', [6].CurrentValue := 1, [6].Mimic := 1, [6].DelayTimer.PRE := 1000, [6].DelayTimerSP := 1, [6].Priority := 1, [6].EnableCfg := 1, [6].ActiveStateCFg := 1, [6].RealInputCfg := 1, [6].InputAddressCfg := 6, [7].Tag := 'XS003', [7].CurrentValue := 1, [7].Mimic := 1, [7].DelayTimer.PRE := 1000, [7].DelayTimerSP := 1, [7].Priority := 1, [7].EnableCfg := 1, [7].ActiveStateCFg := 1, [7].RealInputCfg := 1, [7].InputAddressCfg := 7, [8].Tag := 'SIC001DF', [8].CurrentValue := 1, [8].Mimic := 1, [8].DelayTimer.PRE := 1000, [8].DelayTimerSP := 1, [8].Priority := 1, [8].EnableCfg := 1, [8].ActiveStateCFg := 1, [8].RealInputCfg := 1, [8].InputAddressCfg := 8, [9].Tag := 'SIC002DF', [9].CurrentValue := 1, [9].Mimic := 1, [9].DelayTimer.PRE := 1000, [9].DelayTimerSP := 1, [9].Priority := 1, [9].EnableCfg := 1,
        [9].ActiveStateCFg := 1, [9].RealInputCfg := 1, [9].InputAddressCfg := 9, [10].Tag := 'PSL603', [10].CurrentValue := 1, [10].Mimic := 1, [10].DelayTimer.PRE := 1000, [10].DelayTimerSP := 1, [10].Priority := 1, [10].EnableCfg := 1, [10].ActiveStateCFg := 1, [10].RealInputCfg := 1, [10].InputAddressCfg := 10, [11].Tag := 'XS011', [11].DelayTimerSP := 1, [12].Tag := 'XS012', [12].DelayTimerSP := 1, [13].Tag := 'XC102_3DF', [13].AlarmCurrentValue := 1, [13].DelayTimer.ACC := 4455, [13].DelayTimer.EN := 1, [13].DelayTimer.TT := 1, [13].DelayTimerSP := 1, [14].Tag := 'SIC003DF', [14].DelayTimer.PRE := 2000, [14].DelayTimerSP := 2, [14].EnableCfg := 1, [14].ActiveStateCFg := 1, [14].RealInputCfg := 1, [14].InputAddressCfg := 14, [15].Tag := 'SRL001', [15].SoftInput := 1, [15].DelayTimer.PRE := 2000, [15].DelayTimerSP := 2, [15].EnableCfg := 1, [15].ActiveStateCFg := 1, [15].RealInputCfg := 1, [15].InputAddressCfg := 15, [16].AlarmCurrentValue := 1, [16].Override := 1, [16].SoftInput := 1, [16].DelayTimer.PRE := 1000, [16].DelayTimer.ACC := 1028, [16].DelayTimer.EN := 1, [16].DelayTimer.DN := 1, [16].DelayTimerSP := 1, [16].Priority := 1, [16].EnableCfg := 1, [16].ActiveStateCFg := 1, [16].RealInputCfg := 1, [16].InputAddressCfg := 16, [16].AlarmCfg := 1, [16].OverrideCfg := 1, [16].PriorityCfg := 1, [17].AlarmCurrentValue := 1, [17].Override := 1, [17].SoftInput := 1, [17].DelayTimer.PRE := 1000, [17].DelayTimer.ACC := 1029, [17].DelayTimer.EN := 1,
        [17].DelayTimer.DN := 1, [17].DelayTimerSP := 1, [17].Priority := 1, [17].EnableCfg := 1, [17].ActiveStateCFg := 1, [17].RealInputCfg := 1, [17].InputAddressCfg := 17, [17].AlarmCfg := 1, [17].OverrideCfg := 1, [17].PriorityCfg := 1, [18].AlarmCurrentValue := 1, [18].Override := 1, [18].DelayTimer.PRE := 1000, [18].DelayTimer.ACC := 1029, [18].DelayTimer.EN := 1, [18].DelayTimer.DN := 1, [18].DelayTimerSP := 1, [18].Priority := 1, [18].EnableCfg := 1, [18].ActiveStateCFg := 1, [18].RealInputCfg := 1, [18].InputAddressCfg := 18, [18].AlarmCfg := 1, [18].OverrideCfg := 1, [18].PriorityCfg := 1, [19].CurrentValue := 1, [19].Mimic := 1, [19].DelayTimer.PRE := 1000, [19].DelayTimerSP := 1, [19].Priority := 1, [19].ActiveStateCFg := 1, [19].RealInputCfg := 1, [19].InputAddressCfg := 19, [19].OverrideCfg := 1, [19].PriorityCfg := 1, [20].CurrentValue := 1, [20].Mimic := 1, [20].DelayTimer.PRE := 1000, [20].DelayTimerSP := 1, [20].Priority := 1, [20].ActiveStateCFg := 1, [20].RealInputCfg := 1, [20].InputAddressCfg := 20, [20].OverrideCfg := 1, [20].PriorityCfg := 1, [21].CurrentValue := 1, [21].Override := 1, [21].Mimic := 1, [21].Priority := 1, [21].EnableCfg := 1, [21].ActiveStateCFg := 1, [21].RealInputCfg := 1, [21].InputAddressCfg := 21, [21].AlarmCfg := 1, [21].OverrideCfg := 1, [22].CurrentValue := 1, [22].Override := 1, [22].Mimic := 1, [22].Priority := 1, [22].EnableCfg := 1,
        [22].ActiveStateCFg := 1, [22].RealInputCfg := 1, [22].InputAddressCfg := 22, [22].AlarmCfg := 1, [22].OverrideCfg := 1, [23].AlarmCurrentValue := 1, [23].Override := 1, [23].DelayTimer.PRE := 1000, [23].DelayTimer.ACC := 1029, [23].DelayTimer.EN := 1, [23].DelayTimer.DN := 1, [23].DelayTimerSP := 1, [23].Priority := 1, [23].EnableCfg := 1, [23].ActiveStateCFg := 1, [23].RealInputCfg := 1, [23].InputAddressCfg := 23, [23].AlarmCfg := 1, [23].OverrideCfg := 1, [23].PriorityCfg := 1, [24].AlarmCurrentValue := 1, [24].Override := 1, [24].DelayTimer.PRE := 1000, [24].DelayTimer.ACC := 1029, [24].DelayTimer.EN := 1, [24].DelayTimer.DN := 1, [24].DelayTimerSP := 1, [24].Priority := 1, [24].EnableCfg := 1, [24].ActiveStateCFg := 1, [24].RealInputCfg := 1, [24].InputAddressCfg := 24, [24].AlarmCfg := 1, [24].OverrideCfg := 1, [24].PriorityCfg := 1, [25].AlarmCurrentValue := 1, [25].Override := 1, [25].DelayTimer.PRE := 1000, [25].DelayTimer.ACC := 1030, [25].DelayTimer.EN := 1, [25].DelayTimer.DN := 1, [25].DelayTimerSP := 1, [25].Priority := 1, [25].EnableCfg := 1, [25].ActiveStateCFg := 1, [25].RealInputCfg := 1, [25].InputAddressCfg := 25, [25].AlarmCfg := 1, [25].OverrideCfg := 1, [25].PriorityCfg := 1, [26].AlarmCurrentValue := 1, [26].Override := 1, [26].DelayTimer.PRE := 1000, [26].DelayTimer.ACC := 1030, [26].DelayTimer.EN := 1, [26].DelayTimer.DN := 1, [26].DelayTimerSP := 1, [26].Priority := 1, [26].EnableCfg := 1, [26].ActiveStateCFg := 1,
        [26].RealInputCfg := 1, [26].InputAddressCfg := 26, [26].AlarmCfg := 1, [26].OverrideCfg := 1, [26].PriorityCfg := 1, [27].AlarmCurrentValue := 1, [27].Override := 1, [27].SoftInput := 1, [27].DelayTimer.PRE := 1000, [27].DelayTimer.ACC := 1029, [27].DelayTimer.EN := 1, [27].DelayTimer.DN := 1, [27].DelayTimerSP := 1, [27].Priority := 1, [27].EnableCfg := 1, [27].ActiveStateCFg := 1, [27].RealInputCfg := 1, [27].InputAddressCfg := 27, [27].AlarmCfg := 1, [27].OverrideCfg := 1, [27].PriorityCfg := 1, [28].AlarmCurrentValue := 1, [28].Override := 1, [28].SoftInput := 1, [28].DelayTimer.PRE := 1000, [28].DelayTimer.ACC := 1029, [28].DelayTimer.EN := 1, [28].DelayTimer.DN := 1, [28].DelayTimerSP := 1, [28].EnableCfg := 1, [28].ActiveStateCFg := 1, [28].RealInputCfg := 1, [28].InputAddressCfg := 28, [28].AlarmCfg := 1, [28].OverrideCfg := 1, [28].PriorityCfg := 1, [29].AlarmCurrentValue := 1, [29].Override := 1, [29].SoftInput := 1, [29].DelayTimer.PRE := 1000, [29].DelayTimer.ACC := 1029, [29].DelayTimer.EN := 1, [29].DelayTimer.DN := 1, [29].DelayTimerSP := 1, [29].Priority := 1, [29].EnableCfg := 1, [29].ActiveStateCFg := 1, [29].RealInputCfg := 1, [29].InputAddressCfg := 29, [29].AlarmCfg := 1, [29].OverrideCfg := 1, [29].PriorityCfg := 1, [30].Override := 1, [30].SoftInput := 1, [30].DelayTimer.PRE := 1000, [30].DelayTimerSP := 1, [30].Priority := 1, [30].EnableCfg := 1, [30].ActiveStateCFg := 1, [30].RealInputCfg := 1,
        [30].InputAddressCfg := 30, [30].OverrideCfg := 1, [30].PriorityCfg := 1, [34].SoftInput := 1, [34].EnableCfg := 1, [34].ActiveStateCFg := 1, [34].RealInputCfg := 1, [34].InputAddressCfg := 34, [35].EnableCfg := 1, [35].ActiveStateCFg := 1, [35].RealInputCfg := 1, [35].InputAddressCfg := 35, [36].SoftInput := 1, [36].EnableCfg := 1, [36].ActiveStateCFg := 1, [36].RealInputCfg := 1, [36].InputAddressCfg := 36, [37].EnableCfg := 1, [37].ActiveStateCFg := 1, [37].RealInputCfg := 1, [37].InputAddressCfg := 37, [38].EnableCfg := 1, [38].ActiveStateCFg := 1, [38].RealInputCfg := 1, [38].InputAddressCfg := 38, [39].SoftInput := 1, [39].EnableCfg := 1, [39].ActiveStateCFg := 1, [39].RealInputCfg := 1, [39].InputAddressCfg := 39, [40].EnableCfg := 1, [40].ActiveStateCFg := 1, [40].RealInputCfg := 1, [40].InputAddressCfg := 40, [41].SoftInput := 1, [41].EnableCfg := 1, [41].ActiveStateCFg := 1, [41].RealInputCfg := 1, [41].InputAddressCfg := 41, [50].Tag := 'YA01', [50].AlarmCurrentValue := 1, [50].Override := 1, [50].SoftInput := 1, [50].Condition1 := 1, [50].DelayTimer.PRE := 60000, [50].DelayTimer.ACC := 754, [50].DelayTimer.EN := 1, [50].DelayTimer.TT := 1, [50].DelayTimerSP := 60, [50].EnableCfg := 1, [50].InputAddressCfg := 50, [50].AlarmCfg := 1, [50].AlarmStateCfg := 1, [50].OverrideCfg := 1, [50].PriorityCfg := 1, [50].Cond1Cfg := 1, [51].Tag := 'YA02', [51].CurrentValue := 1, [51].Override := 1, [51].Condition1 := 1,
        [51].DelayTimer.PRE := 60000, [51].DelayTimerSP := 60, [51].EnableCfg := 1, [51].InputAddressCfg := 51, [51].AlarmCfg := 1, [51].AlarmStateCfg := 1, [51].OverrideCfg := 1, [51].PriorityCfg := 1, [51].Cond1Cfg := 1, [52].Tag := 'YA03', [52].AlarmCurrentValue := 1, [52].Override := 1, [52].SoftInput := 1, [52].Condition1 := 1, [52].DelayTimer.PRE := 80000, [52].DelayTimer.ACC := 23271, [52].DelayTimer.EN := 1, [52].DelayTimer.TT := 1, [52].DelayTimerSP := 80, [52].EnableCfg := 1, [52].InputAddressCfg := 52, [52].AlarmCfg := 1, [52].AlarmStateCfg := 1, [52].OverrideCfg := 1, [52].PriorityCfg := 1, [52].Cond1Cfg := 1, [53].Tag := 'YA04', [53].Override := 1, [53].DelayTimer.PRE := 60000, [53].DelayTimerSP := 60, [53].EnableCfg := 1, [53].ActiveStateCFg := 1, [53].InputAddressCfg := 53, [53].AlarmCfg := 1, [53].AlarmStateCfg := 1, [53].OverrideCfg := 1, [53].PriorityCfg := 1, [54].Tag := 'YA05', [54].Override := 1, [54].DelayTimer.PRE := 60000, [54].DelayTimerSP := 60, [54].EnableCfg := 1, [54].ActiveStateCFg := 1, [54].InputAddressCfg := 54, [54].AlarmCfg := 1, [54].AlarmStateCfg := 1, [54].OverrideCfg := 1, [54].PriorityCfg := 1, [55].Tag := 'YA06', [55].Override := 1, [55].DelayTimer.PRE := 5000, [55].DelayTimerSP := 5, [55].Priority := 1, [55].EnableCfg := 1, [55].ActiveStateCFg := 1, [55].InputAddressCfg := 55, [55].AlarmCfg := 1, [55].AlarmStateCfg := 1, [55].OverrideCfg := 1, [55].PriorityCfg := 1,
        [56].Tag := 'YA07', [56].CurrentValue := 1, [56].AlarmCurrentValue := 1, [56].Override := 1, [56].Mimic := 1, [56].SoftInput := 1, [56].DelayTimer.PRE := 2000, [56].DelayTimer.ACC := 2036, [56].DelayTimer.EN := 1, [56].DelayTimer.DN := 1, [56].DelayTimerSP := 2, [56].EnableCfg := 1, [56].ActiveStateCFg := 1, [56].InputAddressCfg := 56, [56].AlarmCfg := 1, [56].AlarmStateCfg := 1, [56].OverrideCfg := 1, [56].PriorityCfg := 1, [57].Tag := 'YA08', [57].Override := 1, [57].DelayTimer.PRE := 5000, [57].DelayTimerSP := 5, [57].Priority := 1, [57].EnableCfg := 1, [57].ActiveStateCFg := 1, [57].InputAddressCfg := 57, [57].AlarmCfg := 1, [57].AlarmStateCfg := 1, [57].OverrideCfg := 1, [57].PriorityCfg := 1, [58].Tag := 'YA09', [58].CurrentValue := 1, [58].AlarmCurrentValue := 1, [58].Override := 1, [58].Mimic := 1, [58].SoftInput := 1, [58].DelayTimer.PRE := 10000, [58].DelayTimer.ACC := 10032, [58].DelayTimer.EN := 1, [58].DelayTimer.DN := 1, [58].DelayTimerSP := 10, [58].EnableCfg := 1, [58].ActiveStateCFg := 1, [58].InputAddressCfg := 58, [58].AlarmCfg := 1, [58].AlarmStateCfg := 1, [58].OverrideCfg := 1, [58].PriorityCfg := 1, [59].Tag := 'YA10', [59].CurrentValue := 1, [59].Mimic := 1, [59].Priority := 1, [59].EnableCfg := 1, [59].InputAddressCfg := 59, [59].AlarmCfg := 1, [59].AlarmStateCfg := 1, [60].Tag := 'YA11', [60].Override := 1, [60].DelayTimer.PRE := 5000, [60].DelayTimerSP := 5,
        [60].EnableCfg := 1, [60].ActiveStateCFg := 1, [60].InputAddressCfg := 60, [60].AlarmCfg := 1, [60].AlarmStateCfg := 1, [60].OverrideCfg := 1, [60].PriorityCfg := 1, [61].Tag := 'YA12', [61].Override := 1, [61].EnableCfg := 1, [61].ActiveStateCFg := 1, [61].InputAddressCfg := 61, [61].AlarmCfg := 1, [61].AlarmStateCfg := 1, [61].OverrideCfg := 1, [61].PriorityCfg := 1, [62].Tag := 'YA13', [62].Override := 1, [62].DelayTimer.PRE := 2000, [62].DelayTimerSP := 2, [62].EnableCfg := 1, [62].ActiveStateCFg := 1, [62].InputAddressCfg := 62, [62].AlarmCfg := 1, [62].AlarmStateCfg := 1, [62].OverrideCfg := 1, [62].PriorityCfg := 1, [63].Tag := 'YA14', [63].CurrentValue := 1, [63].Mimic := 1, [63].DelayTimer.PRE := 60000, [63].DelayTimerSP := 60, [63].EnableCfg := 1, [63].InputAddressCfg := 63, [63].AlarmCfg := 1, [63].AlarmStateCfg := 1, [64].Tag := 'UserNCr1', [64].CurrentValue := 1, [64].Mimic := 1, [64].EnableCfg := 1, [64].InputAddressCfg := 64, [65].Tag := 'UserCr1', [65].CurrentValue := 1, [65].Mimic := 1, [65].Priority := 1, [65].EnableCfg := 1, [65].InputAddressCfg := 65, [66].Tag := 'UserNCr2', [66].CurrentValue := 1, [66].Mimic := 1, [66].EnableCfg := 1, [66].InputAddressCfg := 66, [67].Tag := 'UserCr2', [67].CurrentValue := 1, [67].Mimic := 1, [67].Priority := 1, [67].EnableCfg := 1, [67].InputAddressCfg := 67, [68].Tag := 'ZSDF', [68].Override := 1,
        [68].DelayTimer.PRE := 1000, [68].DelayTimerSP := 1, [68].Priority := 1, [68].EnableCfg := 1, [68].ActiveStateCFg := 1, [68].InputAddressCfg := 68, [68].AlarmCfg := 1, [68].AlarmStateCfg := 1, [68].OverrideCfg := 1, [68].PriorityCfg := 1, [69].Tag := 'YA15', [69].CurrentValue := 1, [69].AlarmCurrentValue := 1, [69].Override := 1, [69].Mimic := 1, [69].SoftInput := 1, [69].DelayTimer.PRE := 5000, [69].DelayTimer.ACC := 5047, [69].DelayTimer.EN := 1, [69].DelayTimer.DN := 1, [69].DelayTimerSP := 5, [69].Priority := 1, [69].EnableCfg := 1, [69].ActiveStateCFg := 1, [69].InputAddressCfg := 69, [69].AlarmCfg := 1, [69].AlarmStateCfg := 1, [69].OverrideCfg := 1, [69].PriorityCfg := 1, [70].Tag := 'YA16', [70].Override := 1, [70].DelayTimerSP := 5, [70].ActiveStateCFg := 1, [70].InputAddressCfg := 70, [70].OverrideCfg := 1, [70].PriorityCfg := 1, [71].Tag := 'YA17', [71].CurrentValue := 1, [71].AlarmCurrentValue := 1, [71].Override := 1, [71].Mimic := 1, [71].SoftInput := 1, [71].DelayTimer.PRE := 5000, [71].DelayTimer.ACC := 5047, [71].DelayTimer.EN := 1, [71].DelayTimer.DN := 1, [71].DelayTimerSP := 5, [71].EnableCfg := 1, [71].ActiveStateCFg := 1, [71].InputAddressCfg := 71, [71].AlarmCfg := 1, [71].AlarmStateCfg := 1, [71].OverrideCfg := 1, [71].PriorityCfg := 1, [72].Tag := 'YA18', [72].Override := 1, [72].DelayTimer.PRE := 2000, [72].DelayTimerSP := 2, [72].EnableCfg := 1, [72].ActiveStateCFg := 1,
        [72].InputAddressCfg := 72, [72].AlarmCfg := 1, [72].AlarmStateCfg := 1, [72].OverrideCfg := 1, [72].PriorityCfg := 1, [73].Tag := 'YA41', [73].Override := 1, [73].EnableCfg := 1, [73].ActiveStateCFg := 1, [73].InputAddressCfg := 73, [73].AlarmCfg := 1, [73].AlarmStateCfg := 1, [73].OverrideCfg := 1, [74].Tag := 'YA20', [74].DelayTimerSP := 2, [75].Tag := 'YA21', [75].CurrentValue := 1, [75].AlarmCurrentValue := 1, [75].AlarmAck := 1, [75].Mimic := 5, [75].SoftInput := 1, [75].DelayTimer.ACC := 2045, [75].DelayTimer.EN := 1, [75].DelayTimer.DN := 1, [75].DelayTimerSP := 5, [75].AlarmONS := 1, [76].Tag := 'YA22', [76].CurrentValue := 1, [76].AlarmCurrentValue := 1, [76].AlarmAck := 1, [76].Mimic := 5, [76].SoftInput := 1, [76].DelayTimer.ACC := 2044, [76].DelayTimer.EN := 1, [76].DelayTimer.DN := 1, [76].DelayTimerSP := 5, [76].AlarmONS := 1, [77].CurrentValue := 1, [77].Mimic := 1, [77].DelayTimerSP := 2, [78].CurrentValue := 1, [78].AlarmCurrentValue := 1, [78].AlarmAck := 1, [78].Mimic := 5, [78].SoftInput := 1, [78].DelayTimer.ACC := 45, [78].DelayTimer.EN := 1, [78].DelayTimer.DN := 1, [78].DelayTimerSP := 2, [78].AlarmONS := 1, [79].CurrentValue := 1, [79].AlarmCurrentValue := 1, [79].Mimic := 1, [79].DelayTimer.ACC := 44, [79].DelayTimer.EN := 1, [79].DelayTimer.DN := 1, [79].DelayTimerSP := 2, [80].CurrentValue := 1, [80].AlarmCurrentValue := 1, [80].Mimic := 1,
        [80].DelayTimer.ACC := 44, [80].DelayTimer.EN := 1, [80].DelayTimer.DN := 1, [80].DelayTimerSP := 2, [81].CurrentValue := 1, [81].AlarmCurrentValue := 1, [81].Mimic := 1, [81].DelayTimer.ACC := 44, [81].DelayTimer.EN := 1, [81].DelayTimer.DN := 1, [81].DelayTimerSP := 2, [82].CurrentValue := 1, [82].AlarmCurrentValue := 1, [82].Mimic := 1, [82].DelayTimer.ACC := 44, [82].DelayTimer.EN := 1, [82].DelayTimer.DN := 1, [82].DelayTimerSP := 2, [83].CurrentValue := 1, [83].AlarmCurrentValue := 1, [83].AlarmAck := 1, [83].Mimic := 5, [83].SoftInput := 1, [83].DelayTimer.ACC := 44, [83].DelayTimer.EN := 1, [83].DelayTimer.DN := 1, [83].DelayTimerSP := 2, [83].AlarmONS := 1, [84].CurrentValue := 1, [84].Mimic := 1, [84].DelayTimerSP := 2, [85].CurrentValue := 1, [85].AlarmCurrentValue := 1, [85].AlarmAck := 1, [85].Mimic := 3, [85].SoftInput := 1, [85].DelayTimer.ACC := 2021, [85].DelayTimer.EN := 1, [85].DelayTimer.DN := 1, [85].DelayTimerSP := 2, [85].AlarmONS := 1, [86].CurrentValue := 1, [86].Mimic := 1, [86].DelayTimerSP := 2, [87].CurrentValue := 1, [87].Mimic := 1, [87].DelayTimerSP := 2, [88].CurrentValue := 1, [88].Mimic := 1, [88].DelayTimerSP := 2, [89].CurrentValue := 1, [89].Mimic := 1, [89].DelayTimerSP := 2, [90].Tag := 'AI101_SIG', [90].CurrentValue := 1, [90].AlarmCurrentValue := 1, [90].Override := 1, [90].Mimic := 1, [90].SoftInput := 1, [90].DelayTimer.PRE := 10000,
        [90].DelayTimer.ACC := 10034, [90].DelayTimer.EN := 1, [90].DelayTimer.DN := 1, [90].DelayTimerSP := 10, [90].EnableCfg := 1, [90].ActiveStateCFg := 1, [90].InputAddressCfg := 90, [90].AlarmCfg := 1, [90].AlarmStateCfg := 1, [90].OverrideCfg := 1, [90].PriorityCfg := 1, [91].Tag := 'AI102_SIG', [91].CurrentValue := 1, [91].AlarmCurrentValue := 1, [91].Override := 1, [91].Mimic := 1, [91].SoftInput := 1, [91].DelayTimer.PRE := 10000, [91].DelayTimer.ACC := 10035, [91].DelayTimer.EN := 1, [91].DelayTimer.DN := 1, [91].DelayTimerSP := 10, [91].EnableCfg := 1, [91].ActiveStateCFg := 1, [91].InputAddressCfg := 91, [91].AlarmCfg := 1, [91].AlarmStateCfg := 1, [91].OverrideCfg := 1, [91].PriorityCfg := 1, [92].Tag := 'AI103_SIG', [92].CurrentValue := 1, [92].AlarmCurrentValue := 1, [92].Override := 1, [92].Mimic := 1, [92].SoftInput := 1, [92].DelayTimer.PRE := 10000, [92].DelayTimer.ACC := 10035, [92].DelayTimer.EN := 1, [92].DelayTimer.DN := 1, [92].DelayTimerSP := 10, [92].EnableCfg := 1, [92].ActiveStateCFg := 1, [92].InputAddressCfg := 92, [92].AlarmCfg := 1, [92].AlarmStateCfg := 1, [92].OverrideCfg := 1, [92].PriorityCfg := 1, [93].Tag := 'FI101_SIG', [93].CurrentValue := 1, [93].AlarmCurrentValue := 1, [93].Override := 1, [93].Mimic := 1, [93].SoftInput := 1, [93].DelayTimer.PRE := 10000, [93].DelayTimer.ACC := 10035, [93].DelayTimer.EN := 1, [93].DelayTimer.DN := 1, [93].DelayTimerSP := 10, [93].EnableCfg := 1, [93].ActiveStateCFg := 1,
        [93].InputAddressCfg := 93, [93].AlarmCfg := 1, [93].AlarmStateCfg := 1, [93].OverrideCfg := 1, [93].PriorityCfg := 1, [94].Tag := 'WI001_SIG', [94].Override := 1, [94].DelayTimer.PRE := 10000, [94].DelayTimerSP := 10, [94].EnableCfg := 1, [94].ActiveStateCFg := 1, [94].InputAddressCfg := 94, [94].AlarmCfg := 1, [94].AlarmStateCfg := 1, [94].OverrideCfg := 1, [94].PriorityCfg := 1, [95].Tag := 'WI101_SIG', [95].CurrentValue := 1, [95].AlarmCurrentValue := 1, [95].Override := 1, [95].Mimic := 1, [95].SoftInput := 1, [95].DelayTimer.PRE := 10000, [95].DelayTimer.ACC := 10034, [95].DelayTimer.EN := 1, [95].DelayTimer.DN := 1, [95].DelayTimerSP := 10, [95].EnableCfg := 1, [95].ActiveStateCFg := 1, [95].InputAddressCfg := 95, [95].AlarmCfg := 1, [95].AlarmStateCfg := 1, [95].OverrideCfg := 1, [95].PriorityCfg := 1, [96].Tag := 'WI102_SIG', [96].CurrentValue := 1, [96].Override := 1, [96].Mimic := 1, [96].SoftInput := 1, [96].DelayTimer.PRE := 10000, [96].DelayTimerSP := 10, [96].EnableCfg := 1, [96].ActiveStateCFg := 1, [96].InputAddressCfg := 96, [96].AlarmStateCfg := 1, [96].OverrideCfg := 1, [96].PriorityCfg := 1, [97].Tag := 'PI001_SIG', [97].CurrentValue := 1, [97].AlarmCurrentValue := 1, [97].Override := 1, [97].Mimic := 1, [97].SoftInput := 1, [97].DelayTimer.PRE := 10000, [97].DelayTimer.ACC := 10035, [97].DelayTimer.EN := 1, [97].DelayTimer.DN := 1, [97].DelayTimerSP := 10, [97].EnableCfg := 1, [97].ActiveStateCFg := 1,
        [97].InputAddressCfg := 97, [97].AlarmCfg := 1, [97].AlarmStateCfg := 1, [97].OverrideCfg := 1, [97].PriorityCfg := 1, [98].Tag := 'PI002_SIG', [98].Override := 1, [98].DelayTimer.PRE := 10000, [98].DelayTimerSP := 10, [98].EnableCfg := 1, [98].ActiveStateCFg := 1, [98].InputAddressCfg := 98, [98].AlarmCfg := 1, [98].AlarmStateCfg := 1, [98].OverrideCfg := 1, [98].PriorityCfg := 1, [99].Tag := 'PI101_SIG', [99].Override := 1, [99].DelayTimer.PRE := 10000, [99].DelayTimerSP := 10, [99].EnableCfg := 1, [99].ActiveStateCFg := 1, [99].InputAddressCfg := 99, [99].AlarmCfg := 1, [99].AlarmStateCfg := 1, [99].OverrideCfg := 1, [99].PriorityCfg := 1, [100].Tag := 'PI401_SIG', [100].Override := 1, [100].DelayTimer.PRE := 10000, [100].DelayTimerSP := 10, [100].EnableCfg := 1, [100].ActiveStateCFg := 1, [100].InputAddressCfg := 100, [100].AlarmCfg := 1, [100].AlarmStateCfg := 1, [100].OverrideCfg := 1, [100].PriorityCfg := 1, [101].Tag := 'TI001_SIG', [101].CurrentValue := 1, [101].AlarmCurrentValue := 1, [101].Override := 1, [101].Mimic := 1, [101].SoftInput := 1, [101].DelayTimer.PRE := 10000, [101].DelayTimer.ACC := 10034, [101].DelayTimer.EN := 1, [101].DelayTimer.DN := 1, [101].DelayTimerSP := 10, [101].EnableCfg := 1, [101].ActiveStateCFg := 1, [101].InputAddressCfg := 101, [101].AlarmCfg := 1, [101].AlarmStateCfg := 1, [101].OverrideCfg := 1, [101].PriorityCfg := 1, [102].Tag := 'PCV001_SIG', [102].Override := 1, [102].DelayTimer.PRE := 10000, [102].DelayTimerSP := 10,
        [102].EnableCfg := 1, [102].ActiveStateCFg := 1, [102].InputAddressCfg := 102, [102].AlarmCfg := 1, [102].AlarmStateCfg := 1, [102].OverrideCfg := 1, [102].PriorityCfg := 1, [103].Tag := 'PCV101_SIG', [103].Override := 1, [103].DelayTimer.PRE := 10000, [103].DelayTimerSP := 10, [103].EnableCfg := 1, [103].ActiveStateCFg := 1, [103].InputAddressCfg := 103, [103].AlarmCfg := 1, [103].AlarmStateCfg := 1, [103].OverrideCfg := 1, [103].PriorityCfg := 1, [104].Tag := 'MIX001_SIG', [104].Override := 1, [104].DelayTimer.PRE := 10000, [104].DelayTimerSP := 10, [104].EnableCfg := 1, [104].ActiveStateCFg := 1, [104].InputAddressCfg := 104, [104].AlarmCfg := 1, [104].AlarmStateCfg := 1, [104].OverrideCfg := 1, [104].PriorityCfg := 1, [105].Tag := 'AI104_SIG', [105].CurrentValue := 1, [105].AlarmCurrentValue := 1, [105].Override := 1, [105].Mimic := 1, [105].SoftInput := 1, [105].DelayTimer.PRE := 10000, [105].DelayTimer.ACC := 10034, [105].DelayTimer.EN := 1, [105].DelayTimer.DN := 1, [105].DelayTimerSP := 10, [105].EnableCfg := 1, [105].ActiveStateCFg := 1, [105].InputAddressCfg := 105, [105].AlarmCfg := 1, [105].AlarmStateCfg := 1, [105].OverrideCfg := 1, [105].PriorityCfg := 1, [106].CurrentValue := 1, [106].AlarmCurrentValue := 1, [106].Override := 1, [106].Mimic := 1, [106].SoftInput := 1, [106].DelayTimer.PRE := 10000, [106].DelayTimer.ACC := 10034, [106].DelayTimer.EN := 1, [106].DelayTimer.DN := 1, [106].DelayTimerSP := 10, [106].EnableCfg := 1, [106].ActiveStateCFg := 1, [106].InputAddressCfg := 106,
        [106].AlarmCfg := 1, [106].AlarmStateCfg := 1, [106].OverrideCfg := 1, [106].PriorityCfg := 1, [107].CurrentValue := 1, [107].AlarmCurrentValue := 1, [107].AlarmAck := 1, [107].Mimic := 3, [107].SoftInput := 1, [107].DelayTimer.PRE := 10000, [107].DelayTimer.ACC := 41, [107].DelayTimer.EN := 1, [107].DelayTimer.DN := 1, [107].DelayTimerSP := 10, [107].ActiveStateCFg := 1, [107].InputAddressCfg := 107, [107].AlarmStateCfg := 1, [107].OverrideCfg := 1, [107].PriorityCfg := 1, [107].AlarmONS := 1, [108].CurrentValue := 1, [108].Override := 1, [108].Mimic := 1, [108].SoftInput := 1, [108].DelayTimer.PRE := 10000, [108].DelayTimerSP := 10, [108].EnableCfg := 1, [108].ActiveStateCFg := 1, [108].InputAddressCfg := 108, [108].AlarmStateCfg := 1, [108].OverrideCfg := 1, [108].PriorityCfg := 1, [109].CurrentValue := 1, [109].AlarmCurrentValue := 1, [109].Override := 1, [109].Mimic := 1, [109].SoftInput := 1, [109].DelayTimer.PRE := 10000, [109].DelayTimer.ACC := 10035, [109].DelayTimer.EN := 1, [109].DelayTimer.DN := 1, [109].DelayTimerSP := 10, [109].EnableCfg := 1, [109].ActiveStateCFg := 1, [109].InputAddressCfg := 109, [109].AlarmCfg := 1, [109].AlarmStateCfg := 1, [109].OverrideCfg := 1, [109].PriorityCfg := 1, [110].Override := 1, [110].DelayTimer.PRE := 10000, [110].DelayTimerSP := 10, [110].EnableCfg := 1, [110].ActiveStateCFg := 1, [110].InputAddressCfg := 110, [110].AlarmCfg := 1, [110].AlarmStateCfg := 1, [110].OverrideCfg := 1, [110].PriorityCfg := 1, [111].CurrentValue := 1,
        [111].AlarmCurrentValue := 1, [111].Override := 1, [111].Mimic := 1, [111].SoftInput := 1, [111].DelayTimer.PRE := 10000, [111].DelayTimer.ACC := 10032, [111].DelayTimer.EN := 1, [111].DelayTimer.DN := 1, [111].DelayTimerSP := 10, [111].EnableCfg := 1, [111].ActiveStateCFg := 1, [111].InputAddressCfg := 111, [111].AlarmCfg := 1, [111].AlarmStateCfg := 1, [111].OverrideCfg := 1, [111].PriorityCfg := 1);   // Digital Point Array
        [110]   // Retentate Flow Signal default
        [111]   // Filtrate Temperature Signal Default
        [54]   // Database Overload
        [30]   // TCU Defect
        [14]   // Pump P001 Type
        [34]   // Exchange DI#1
        [21]   // Feed Pump High Pressure
        [0]   // Valves Air Defect
        [100]   // Transfer Pump Pressure Signal Default
        [101]   // Feed Tank Temperature Signal Default
        [102]   // PCV101 Position Signal Default
        [103]   // PCV201 Position Signal Default
        [104]   // Mixer Speed Signal Default
        [105]   // Filtrate pH Signal Default
        [106]   // Feed Tank pH Signal default
        [107]   // Feed Tank Conductivity Signal default
        [108]   // TCU Temperature Signal default
        [109]   // Filtrate Conductivity Cleaning Signal default
        [10]   // Clamshell Locking 5 Closed
        [50]   // PC to PLC communication failure
        [15]   // Pump P002 Type
        [19]   // H100 pH Defect
        [16]   // P001 Defect
        [17]   // P002 Defect
        [18]   // C8000 Defect
        [1]   // Manifold Valves Air Defect
        [20]   // H100 Cond Defect
        [25]   // Pump Cart 24 VDC Defect
        [22]   // Transfer Pump High Pressure
        [23]   // P001 48 VDC Defect
        [24]   // P002 48 VDC Defect
        [59]   // PLC Program Major Fault
        [27]   // Pump P003 Power Supply Defect
        [28]   // Mixer Defect
        [29]   // P003 Defect
        [2]   // Emergency Stop
        [3]   // Reset Buzzer
        [35]   // Exchange DI#2
        [36]   // Exchange DI#3
        [37]   // Exchange DI#4
        [38]   // Exchange DI#5
        [39]   // Exchange DI#6
        [40]   // Exchange DI#7
        [41]   // Exchange DI#8
        [4]   // 24 VDC defect
        [98]   // Rentate Pressure Signal Default
        [51]   // CCP Runtime communication failure
        [52]   // Historical Data collection failure
        [55]   // Node 0 communication failure
        [56]   // Node 0 internal defect
        [57]   // Node 1 communication failure
        [58]   // Node 1 internal defect
        [73]   // Operating Time Exceeded
        [5]   // Door Closed
        [60]   // Database Corrupted
        [61]   // Unauthorized Accesses
        [62]   // Tank Size Mismatch
        [63]   // SQL Server Write Failure
        [64]   // User Non Critical Alarm 1
        [65]   // User Critical Alarm 1
        [66]   // User Non Critical Alarm 2
        [67]   // User Critical Alarm 2
        [68]   // ZSDF Clamshell Locking Defect
        [69]   // ACT350 Communication Failure
        [6]   // Clamshell Locking 1 Closed
        [70]   // Watchdog Gateway
        [71]   // Mobius Device Communication Failure
        [72]   // Pump Type Mismatch
        [7]   // Clamshell Locking 2 Closed
        [8]   // Clamshell Locking 3 Closed
        [90]   // Filtrate Conductivity Process Signal default
        [91]   // Filtrate UV1 Signal default
        [92]   // Filtrate UV2 Signal default
        [93]   // Filtrate Flow Signal default
        [94]   // Transfer Pump Flow Signal default
        [95]   // Feed Tank Pressure Signal default
        [96]   // External Filtrate Weight Signal default
        [97]   // Feed Pressure Signal Default
        [99]   // Filtrate Pressure Signal Default
        [9]   // Clamshell Locking 4 Closed
        [26]   // Mixer 48 VDC Defect
        [53]   // Hard Drive Overload
   DigitalPoint_Storage : DigitalPoint[6,150] := ([0,0].Tag := 'PISL601', [0,0].AlarmCurrentValue := 1, [0,0].AlarmAck := 1, [0,0].Alarm := 1, [0,0].Mimic := 5, [0,0].DelayTimer.PRE := 2000, [0,0].DelayTimer.ACC := 2025, [0,0].DelayTimer.EN := 1, [0,0].DelayTimer.DN := 1, [0,0].DelayTimerSP := 2, [0,0].Priority := 1, [0,0].EnableCfg := 1, [0,0].ActiveStateCFg := 1, [0,0].RealInputCfg := 1, [0,0].AlarmCfg := 1, [0,0].OverrideCfg := 1, [0,0].PriorityCfg := 1, [0,0].AlarmONS := 1, [0,1].Tag := 'PISL602', [0,1].AlarmCurrentValue := 1, [0,1].AlarmAck := 1, [0,1].Alarm := 1, [0,1].Mimic := 5, [0,1].Condition2 := 1, [0,1].DelayTimer.PRE := 2000, [0,1].DelayTimer.ACC := 2053, [0,1].DelayTimer.EN := 1, [0,1].DelayTimer.DN := 1, [0,1].DelayTimerSP := 2, [0,1].Priority := 1, [0,1].EnableCfg := 1, [0,1].ActiveStateCFg := 1, [0,1].RealInputCfg := 1, [0,1].InputAddressCfg := 1, [0,1].AlarmCfg := 1, [0,1].OverrideCfg := 1, [0,1].PriorityCfg := 1, [0,1].AlarmONS := 1, [0,2].Tag := 'ES001', [0,2].AlarmCurrentValue := 1, [0,2].AlarmAck := 1, [0,2].Alarm := 1, [0,2].Mimic := 5, [0,2].DelayTimer.PRE := 1000, [0,2].DelayTimer.ACC := 1047, [0,2].DelayTimer.EN := 1, [0,2].DelayTimer.DN := 1, [0,2].DelayTimerSP := 1, [0,2].Priority := 1, [0,2].EnableCfg := 1, [0,2].ActiveStateCFg := 1, [0,2].RealInputCfg := 1, [0,2].InputAddressCfg := 2, [0,2].AlarmCfg := 1, [0,2].AlarmONS := 1, [0,3].Tag := 'RSBUZZ', [0,3].DelayTimer.PRE := 2000, [0,3].DelayTimerSP := 2, [0,3].EnableCfg := 1, [0,3].ActiveStateCFg := 1,
        [0,3].RealInputCfg := 1, [0,3].InputAddressCfg := 3, [0,4].Tag := 'DF24VDC', [0,4].AlarmCurrentValue := 1, [0,4].AlarmAck := 1, [0,4].Alarm := 1, [0,4].Mimic := 5, [0,4].DelayTimer.PRE := 1000, [0,4].DelayTimer.ACC := 1048, [0,4].DelayTimer.EN := 1, [0,4].DelayTimer.DN := 1, [0,4].DelayTimerSP := 1, [0,4].Priority := 1, [0,4].EnableCfg := 1, [0,4].ActiveStateCFg := 1, [0,4].RealInputCfg := 1, [0,4].InputAddressCfg := 4, [0,4].AlarmCfg := 1, [0,4].OverrideCfg := 1, [0,4].PriorityCfg := 1, [0,4].AlarmONS := 1, [0,5].Tag := 'ZS008', [0,5].AlarmCurrentValue := 1, [0,5].AlarmAck := 1, [0,5].Alarm := 1, [0,5].Mimic := 5, [0,5].DelayTimer.PRE := 1000, [0,5].DelayTimer.ACC := 1048, [0,5].DelayTimer.EN := 1, [0,5].DelayTimer.DN := 1, [0,5].DelayTimerSP := 1, [0,5].Priority := 1, [0,5].EnableCfg := 1, [0,5].ActiveStateCFg := 1, [0,5].RealInputCfg := 1, [0,5].InputAddressCfg := 5, [0,5].AlarmCfg := 1, [0,5].OverrideCfg := 1, [0,5].AlarmONS := 1, [0,6].Tag := 'ZS001', [0,6].DelayTimer.PRE := 2000, [0,6].DelayTimerSP := 2, [0,6].EnableCfg := 1, [0,6].ActiveStateCFg := 1, [0,6].RealInputCfg := 1, [0,6].InputAddressCfg := 6, [0,7].Tag := 'ZS002', [0,7].DelayTimer.PRE := 2000, [0,7].DelayTimerSP := 2, [0,7].EnableCfg := 1, [0,7].ActiveStateCFg := 1, [0,7].RealInputCfg := 1, [0,7].InputAddressCfg := 7, [0,8].Tag := 'ZS003', [0,8].DelayTimer.PRE := 2000, [0,8].DelayTimerSP := 2, [0,8].EnableCfg := 1, [0,8].ActiveStateCFg := 1, [0,8].RealInputCfg := 1, [0,8].InputAddressCfg := 8,
        [0,9].Tag := 'ZS004', [0,9].DelayTimer.PRE := 2000, [0,9].DelayTimerSP := 2, [0,9].EnableCfg := 1, [0,9].ActiveStateCFg := 1, [0,9].RealInputCfg := 1, [0,9].InputAddressCfg := 9, [0,10].Tag := 'ZS005', [0,10].DelayTimer.PRE := 2000, [0,10].DelayTimerSP := 2, [0,10].EnableCfg := 1, [0,10].ActiveStateCFg := 1, [0,10].RealInputCfg := 1, [0,10].InputAddressCfg := 10, [0,11].Tag := 'ZS006', [0,11].DelayTimer.PRE := 2000, [0,11].DelayTimerSP := 2, [0,11].EnableCfg := 1, [0,11].ActiveStateCFg := 1, [0,11].RealInputCfg := 1, [0,11].InputAddressCfg := 11, [0,12].Tag := 'ZS007', [0,12].DelayTimer.PRE := 2000, [0,12].DelayTimerSP := 2, [0,12].EnableCfg := 1, [0,12].ActiveStateCFg := 1, [0,12].RealInputCfg := 1, [0,12].InputAddressCfg := 12, [0,13].Tag := 'ZS008', [0,13].AlarmCurrentValue := 1, [0,13].DelayTimer.PRE := 20000, [0,13].DelayTimerSP := 2, [0,13].Priority := 1, [0,13].EnableCfg := 1, [0,13].ActiveStateCFg := 1, [0,13].RealInputCfg := 1, [0,13].InputAddressCfg := 13, [0,13].AlarmCfg := 1, [0,13].OverrideCfg := 1, [0,13].PriorityCfg := 1, [0,13].Cond1Cfg := 1, [0,14].Tag := 'XS011', [0,14].DelayTimer.PRE := 2000, [0,14].DelayTimerSP := 2, [0,14].EnableCfg := 1, [0,14].ActiveStateCFg := 1, [0,14].RealInputCfg := 1, [0,14].InputAddressCfg := 14, [0,15].Tag := 'XS012', [0,15].SoftInput := 1, [0,15].DelayTimer.PRE := 2000, [0,15].DelayTimerSP := 2, [0,15].EnableCfg := 1, [0,15].ActiveStateCFg := 1, [0,15].RealInputCfg := 1, [0,15].InputAddressCfg := 15, [0,16].Tag := 'SIC001DF', [0,16].AlarmCurrentValue := 1, [0,16].AlarmAck := 1, [0,16].Alarm := 1,
        [0,16].Mimic := 5, [0,16].SoftInput := 1, [0,16].DelayTimer.PRE := 1000, [0,16].DelayTimer.ACC := 1046, [0,16].DelayTimer.EN := 1, [0,16].DelayTimer.DN := 1, [0,16].DelayTimerSP := 1, [0,16].Priority := 1, [0,16].EnableCfg := 1, [0,16].ActiveStateCFg := 1, [0,16].RealInputCfg := 1, [0,16].InputAddressCfg := 16, [0,16].AlarmCfg := 1, [0,16].OverrideCfg := 1, [0,16].PriorityCfg := 1, [0,16].AlarmONS := 1, [0,17].Tag := 'SIC002DF', [0,17].AlarmCurrentValue := 1, [0,17].AlarmAck := 1, [0,17].Alarm := 1, [0,17].Mimic := 5, [0,17].SoftInput := 1, [0,17].DelayTimer.PRE := 1000, [0,17].DelayTimer.ACC := 1046, [0,17].DelayTimer.EN := 1, [0,17].DelayTimer.DN := 1, [0,17].DelayTimerSP := 1, [0,17].Priority := 1, [0,17].EnableCfg := 1, [0,17].ActiveStateCFg := 1, [0,17].RealInputCfg := 1, [0,17].InputAddressCfg := 17, [0,17].AlarmCfg := 1, [0,17].OverrideCfg := 1, [0,17].PriorityCfg := 1, [0,17].AlarmONS := 1, [0,18].Tag := 'AA008', [0,18].AlarmCurrentValue := 1, [0,18].AlarmAck := 1, [0,18].Alarm := 1, [0,18].Mimic := 5, [0,18].DelayTimer.PRE := 1000, [0,18].DelayTimer.ACC := 1046, [0,18].DelayTimer.EN := 1, [0,18].DelayTimer.DN := 1, [0,18].DelayTimerSP := 1, [0,18].Priority := 1, [0,18].EnableCfg := 1, [0,18].ActiveStateCFg := 1, [0,18].RealInputCfg := 1, [0,18].InputAddressCfg := 18, [0,18].AlarmCfg := 1, [0,18].OverrideCfg := 1, [0,18].PriorityCfg := 1, [0,18].AlarmONS := 1, [0,19].Tag := 'LSH001', [0,19].AlarmCurrentValue := 1, [0,19].Override := 1, [0,19].DelayTimer.PRE := 1000, [0,19].DelayTimer.ACC := 1058,
        [0,19].DelayTimer.EN := 1, [0,19].DelayTimer.DN := 1, [0,19].DelayTimerSP := 1, [0,19].EnableCfg := 1, [0,19].ActiveStateCFg := 1, [0,19].RealInputCfg := 1, [0,19].InputAddressCfg := 19, [0,19].AlarmCfg := 1, [0,19].OverrideCfg := 1, [0,19].PriorityCfg := 1, [0,20].Tag := 'LSL002', [0,20].AlarmCurrentValue := 1, [0,20].Override := 1, [0,20].DelayTimer.PRE := 1000, [0,20].DelayTimer.ACC := 1059, [0,20].DelayTimer.EN := 1, [0,20].DelayTimer.DN := 1, [0,20].DelayTimerSP := 1, [0,20].EnableCfg := 1, [0,20].ActiveStateCFg := 1, [0,20].RealInputCfg := 1, [0,20].InputAddressCfg := 20, [0,20].AlarmCfg := 1, [0,20].OverrideCfg := 1, [0,20].PriorityCfg := 1, [0,21].Tag := 'PSH001', [0,21].AlarmCurrentValue := 1, [0,21].AlarmAck := 1, [0,21].Alarm := 1, [0,21].Mimic := 5, [0,21].DelayTimer.PRE := 1000, [0,21].DelayTimer.ACC := 1045, [0,21].DelayTimer.EN := 1, [0,21].DelayTimer.DN := 1, [0,21].DelayTimerSP := 1, [0,21].Priority := 1, [0,21].EnableCfg := 1, [0,21].ActiveStateCFg := 1, [0,21].RealInputCfg := 1, [0,21].InputAddressCfg := 21, [0,21].AlarmCfg := 1, [0,21].AlarmONS := 1, [0,22].Tag := 'PSH002', [0,22].AlarmCurrentValue := 1, [0,22].AlarmAck := 1, [0,22].Alarm := 1, [0,22].Mimic := 5, [0,22].DelayTimer.PRE := 1000, [0,22].DelayTimer.ACC := 1045, [0,22].DelayTimer.EN := 1, [0,22].DelayTimer.DN := 1, [0,22].DelayTimerSP := 1, [0,22].Priority := 1, [0,22].EnableCfg := 1, [0,22].ActiveStateCFg := 1, [0,22].RealInputCfg := 1, [0,22].InputAddressCfg := 22, [0,22].AlarmCfg := 1, [0,22].AlarmONS := 1, [0,23].Tag := 'DF48VP001',
        [0,23].AlarmCurrentValue := 1, [0,23].AlarmAck := 1, [0,23].Alarm := 1, [0,23].Mimic := 5, [0,23].DelayTimer.PRE := 1000, [0,23].DelayTimer.ACC := 1045, [0,23].DelayTimer.EN := 1, [0,23].DelayTimer.DN := 1, [0,23].DelayTimerSP := 1, [0,23].Priority := 1, [0,23].EnableCfg := 1, [0,23].ActiveStateCFg := 1, [0,23].RealInputCfg := 1, [0,23].InputAddressCfg := 23, [0,23].AlarmCfg := 1, [0,23].OverrideCfg := 1, [0,23].PriorityCfg := 1, [0,23].AlarmONS := 1, [0,24].Tag := 'DF48VP002', [0,24].AlarmCurrentValue := 1, [0,24].AlarmAck := 1, [0,24].Alarm := 1, [0,24].Mimic := 5, [0,24].DelayTimer.PRE := 1000, [0,24].DelayTimer.ACC := 1046, [0,24].DelayTimer.EN := 1, [0,24].DelayTimer.DN := 1, [0,24].DelayTimerSP := 1, [0,24].Priority := 1, [0,24].EnableCfg := 1, [0,24].ActiveStateCFg := 1, [0,24].RealInputCfg := 1, [0,24].InputAddressCfg := 24, [0,24].AlarmCfg := 1, [0,24].OverrideCfg := 1, [0,24].PriorityCfg := 1, [0,24].AlarmONS := 1, [0,25].Tag := 'XS002', [0,25].AlarmCurrentValue := 1, [0,25].DelayTimer.PRE := 20000, [0,25].DelayTimerSP := 2, [0,25].Priority := 1, [0,25].EnableCfg := 1, [0,25].ActiveStateCFg := 1, [0,25].RealInputCfg := 1, [0,25].InputAddressCfg := 25, [0,25].AlarmCfg := 1, [0,25].OverrideCfg := 1, [0,25].PriorityCfg := 1, [0,25].Cond1Cfg := 1, [0,26].Override := 1, [0,26].ActiveStateCFg := 1, [0,26].RealInputCfg := 1, [0,26].InputAddressCfg := 26, [0,26].OverrideCfg := 1, [0,26].PriorityCfg := 1, [0,27].Override := 1, [0,27].SoftInput := 1, [0,27].ActiveStateCFg := 1, [0,27].RealInputCfg := 1,
        [0,27].InputAddressCfg := 27, [0,27].OverrideCfg := 1, [0,27].PriorityCfg := 1, [0,28].Override := 1, [0,28].SoftInput := 1, [0,28].ActiveStateCFg := 1, [0,28].RealInputCfg := 1, [0,28].InputAddressCfg := 28, [0,28].OverrideCfg := 1, [0,28].PriorityCfg := 1, [0,29].Override := 1, [0,29].SoftInput := 1, [0,29].ActiveStateCFg := 1, [0,29].RealInputCfg := 1, [0,29].InputAddressCfg := 29, [0,29].OverrideCfg := 1, [0,29].PriorityCfg := 1, [0,30].Override := 1, [0,30].SoftInput := 1, [0,30].ActiveStateCFg := 1, [0,30].RealInputCfg := 1, [0,30].InputAddressCfg := 30, [0,30].OverrideCfg := 1, [0,30].PriorityCfg := 1, [0,31].Override := 1, [0,31].ActiveStateCFg := 1, [0,31].RealInputCfg := 1, [0,31].InputAddressCfg := 31, [0,31].OverrideCfg := 1, [0,31].PriorityCfg := 1, [0,34].Tag := 'DI1', [0,34].Override := 1, [0,34].SoftInput := 1, [0,34].EnableCfg := 1, [0,34].ActiveStateCFg := 1, [0,34].RealInputCfg := 1, [0,34].InputAddressCfg := 34, [0,34].OverrideCfg := 1, [0,34].PriorityCfg := 1, [0,35].Tag := 'DI2', [0,35].Override := 1, [0,35].EnableCfg := 1, [0,35].ActiveStateCFg := 1, [0,35].RealInputCfg := 1, [0,35].InputAddressCfg := 35, [0,35].OverrideCfg := 1, [0,35].PriorityCfg := 1, [0,36].Tag := 'DI3', [0,36].Override := 1, [0,36].SoftInput := 1, [0,36].EnableCfg := 1, [0,36].ActiveStateCFg := 1, [0,36].RealInputCfg := 1, [0,36].InputAddressCfg := 36, [0,36].OverrideCfg := 1, [0,36].PriorityCfg := 1, [0,37].Tag := 'DI4', [0,37].Override := 1, [0,37].EnableCfg := 1, [0,37].ActiveStateCFg := 1,
        [0,37].RealInputCfg := 1, [0,37].InputAddressCfg := 37, [0,37].OverrideCfg := 1, [0,37].PriorityCfg := 1, [0,38].Tag := 'DI5', [0,38].Override := 1, [0,38].EnableCfg := 1, [0,38].ActiveStateCFg := 1, [0,38].RealInputCfg := 1, [0,38].InputAddressCfg := 38, [0,38].OverrideCfg := 1, [0,38].PriorityCfg := 1, [0,39].Tag := 'DI6', [0,39].Override := 1, [0,39].SoftInput := 1, [0,39].EnableCfg := 1, [0,39].ActiveStateCFg := 1, [0,39].RealInputCfg := 1, [0,39].InputAddressCfg := 39, [0,39].OverrideCfg := 1, [0,39].PriorityCfg := 1, [0,40].Tag := 'DI7', [0,40].Override := 1, [0,40].EnableCfg := 1, [0,40].ActiveStateCFg := 1, [0,40].RealInputCfg := 1, [0,40].InputAddressCfg := 40, [0,40].OverrideCfg := 1, [0,40].PriorityCfg := 1, [0,41].Tag := 'DI8', [0,41].Override := 1, [0,41].EnableCfg := 1, [0,41].ActiveStateCFg := 1, [0,41].RealInputCfg := 1, [0,41].InputAddressCfg := 41, [0,41].OverrideCfg := 1, [0,41].PriorityCfg := 1, [0,50].Tag := 'YA01', [0,50].Desc := 'PC to PLC Com. Failure', [0,50].AlarmCurrentValue := 1, [0,50].SoftInput := 1, [0,50].Condition1 := 1, [0,50].Cond1Text := 'HMI HeartBeat received', [0,50].DelayTimer.PRE := 60000, [0,50].DelayTimer.ACC := 442, [0,50].DelayTimer.EN := 1, [0,50].DelayTimer.TT := 1, [0,50].DelayTimerSP := 60, [0,50].EnableCfg := 1, [0,50].InputAddressCfg := 50, [0,50].AlarmCfg := 1, [0,50].AlarmStateCfg := 1, [0,50].OverrideCfg := 1, [0,50].PriorityCfg := 1, [0,50].Cond1Cfg := 1, [0,51].Tag := 'YA02', [0,51].Desc := 'CCP Runtime Com. Failure', [0,51].AlarmCurrentValue := 1, [0,51].Alarm := 1, [0,51].Mimic := 2,
        [0,51].SoftInput := 1, [0,51].Condition1 := 1, [0,51].Cond1Text := 'HMI HeartBeat received', [0,51].DelayTimer.PRE := 60000, [0,51].DelayTimer.ACC := 60061, [0,51].DelayTimer.EN := 1, [0,51].DelayTimer.DN := 1, [0,51].DelayTimerSP := 60, [0,51].EnableCfg := 1, [0,51].InputAddressCfg := 51, [0,51].AlarmCfg := 1, [0,51].AlarmStateCfg := 1, [0,51].OverrideCfg := 1, [0,51].PriorityCfg := 1, [0,51].Cond1Cfg := 1, [0,51].AlarmONS := 1, [0,52].Tag := 'YA03', [0,52].Desc := 'Hist. Data Collect. Fail', [0,52].AlarmCurrentValue := 1, [0,52].Alarm := 1, [0,52].Mimic := 2, [0,52].SoftInput := 1, [0,52].Condition1 := 1, [0,52].Cond1Text := 'HMI HeartBeat received', [0,52].DelayTimer.PRE := 60000, [0,52].DelayTimer.ACC := 1286, [0,52].DelayTimer.EN := 1, [0,52].DelayTimer.TT := 1, [0,52].DelayTimerSP := 60, [0,52].EnableCfg := 1, [0,52].InputAddressCfg := 52, [0,52].AlarmCfg := 1, [0,52].AlarmStateCfg := 1, [0,52].OverrideCfg := 1, [0,52].PriorityCfg := 1, [0,52].Cond1Cfg := 1, [0,52].AlarmONS := 1, [0,53].Tag := 'YA04', [0,53].Desc := 'HDD OverLoad', [0,53].DelayTimer.PRE := 60000, [0,53].DelayTimerSP := 60, [0,53].EnableCfg := 1, [0,53].ActiveStateCFg := 1, [0,53].InputAddressCfg := 53, [0,53].AlarmCfg := 1, [0,53].AlarmStateCfg := 1, [0,53].OverrideCfg := 1, [0,53].PriorityCfg := 1, [0,54].Tag := 'YA05', [0,54].DelayTimer.PRE := 60000, [0,54].DelayTimerSP := 60, [0,54].EnableCfg := 1, [0,54].ActiveStateCFg := 1, [0,54].InputAddressCfg := 54, [0,54].AlarmCfg := 1, [0,54].AlarmStateCfg := 1, [0,54].OverrideCfg := 1, [0,54].PriorityCfg := 1, [0,55].Tag := 'YA06', [0,55].CurrentValue := 1,
